(* IEC 61131-3 sources: JingjiangArm/moonboxpro_arm_8.4/Application/Application/任务列表/ExtTask/动作处理/预套准, 13 files *)

(* ---- ENUM_MotionStepIDs.st ---- *)
(*@CES
Name=ENUM_MotionStepIDs
Type=Gvl
TypeGuid=2db5746d-d284-4425-9f7f-2663a34b0ebc
Guid=2f95a26a-5938-4297-8364-5fa39176fcfb
HasDeclaration=True
HasImplementation=False
*)
{DECLARATION}

TYPE ENUM_MotionStepIDs : (
	MOTION_STEP_NothingDo						:= -1,(*啥都不做*)
	MOTION_STEP_MotionCtrlModel				:= 9,(*2021.2.21.134018设置运动模式设置|+Liu.yt*)
	MOTION_STEP_ServoOff					:= 10,(*下伺服|*)
	MOTION_STEP_ClrSts						:= 11,(*清错误状态|*)
	MOTION_STEP_ZeroPos						:= 12,(*清位置|*)
	MOTION_STEP_ZeroPos_Again				:= 13,(*2018.9.4.144137\再次清位置|*)
	MOTION_STEP_ServoOn						:= 14,(*上伺服|*)
	MOTION_STEP_PtModeDynamic				:= 15,(*设置动态pt规划|*)
	MOTION_STEP_PtClear						:= 16,(*清除动态ptFIFO|*)
	MOTION_STEP_SetModal0					:= 17,(*2017-09-11 09:14:16| 模态0*)
	MOTION_STEP_SyncAllModal0				:= 18,(*同步所有轴模态|*)
	MOTION_STEP_SetModal1					:= 19,(*2017-09-11 09:14:24| 模态1*)
	MOTION_STEP_SyncAllModal1				:= 20,(*同步所有轴模态|*)
	MOTION_STEP_WaitingModalChanged			:= 21,(*等待模态切换0到1|*)
	MOTION_STEP_PushInitialPTdata			:= 22,(*压入初始的几段PT数据*)
	MOTION_STEP_WritePT						:= 23,(*写pt*)
	MOTION_STEP_CheckPTPrf					:= 24,(*检查pt规划器*)
	MOTION_STEP_SetTpid						:= 25,(*设置前馈增益|*)
	MOTION_STEP_SetPosErr					:= 26,(*设置位置偏差|*)
	MOTION_STEP_SetEncSns					:= 27,(*编码器反转|*)
	MOTION_STEP_CheckAllServoSts			:= 28,(*检查所有上伺服的状态|*)
	MOTION_STEP_WillLeaveWritePT			:= 29,(*将要离开PT写操作|2019.11.29.143804_*)
	MOTION_STEP_MULTI_GTCMD					:= 30,(*多个指令同时执行标志@单运行功能使用|点了按钮响应太慢了*)
	MOTION_STEP_ErrorOccured				:= 110(*错误发生*)
);
END_TYPE
{IMPLEMENTATION}

(* ---- KS_CalcCircleTangentDistance.st ---- *)
(*@CES
Name=KS_CalcCircleTangentDistance
Type=FunctionBlock
TypeGuid=6f9dac99-8de1-4efc-8465-68ac443b7d08
Guid=1060efe6-291c-4829-ad87-f7b1dbfd88c0
HasDeclaration=True
HasImplementation=True
*)
{DECLARATION}
FUNCTION KS_CalcCircleTangentDistance : LREAL(*计算两个圆的切线距离|*)
VAR_INPUT
	i_lrX_Circle0							: LREAL;(*圆1的圆心坐标x|*)
	i_lrY_Circle0							: LREAL;(*圆1的圆心坐标y|*)
	i_lrDiam_Circle0						: LREAL;(*圆1的直径|*)
	i_lrX_Circle1							: LREAL;(*圆2的圆心坐标x|*)
	i_lrY_Circle1							: LREAL;(*圆2的圆心坐标y|*)
	i_lrDiam_Circle1						: LREAL;(*圆2的直径|*)
	i_xAtSameSide							: BOOL;(*TRUE表示圆是在切线的同一边(外公切)|FALSE表示分别在切线的两边(内公切)|*)
END_VAR
VAR
	lrN										: LREAL;
	lrResult								: LREAL;
	lrCenterDistance						: LREAL;(*两个圆的圆心距|*)
END_VAR
{IMPLEMENTATION}
lrResult:= 0;

(*
/.圆心距|
/.直角三角形的斜边|
/.*)
lrCenterDistance:= SQRT((i_lrX_Circle0-i_lrX_Circle1)*(i_lrX_Circle0-i_lrX_Circle1)+(i_lrY_Circle0-i_lrY_Circle1)*(i_lrY_Circle0-i_lrY_Circle1));
IF i_xAtSameSide THEN
	(*
	/.外公切|
	/.外公切线的长=根号下[圆心距的平方-（大圆半径减小圆半径）的平方]|
	/.*)
	lrN:= (lrCenterDistance*lrCenterDistance)-(((i_lrDiam_Circle0-i_lrDiam_Circle1)/2)*((i_lrDiam_Circle0-i_lrDiam_Circle1)/2));
	IF lrN<0 THEN
		;
	ELSE
		lrResult:= SQRT(lrN);
	END_IF
ELSE
	(*
	/.内公切|
	/.内公切线的长=根号下[圆心距的平方-（大圆半径加小圆半径）的平方]|
	/.*)
	lrN:= (lrCenterDistance*lrCenterDistance)-(((i_lrDiam_Circle0+i_lrDiam_Circle1)/2)*((i_lrDiam_Circle0+i_lrDiam_Circle1)/2));
	IF lrN<0 THEN
		;
	ELSE
		lrResult:= SQRT(lrN);
	END_IF
END_IF
KS_CalcCircleTangentDistance:= lrResult;

(* ---- KS_CalcForPreRegister.st ---- *)
(*@CES
Name=KS_CalcForPreRegister
Type=FunctionBlock
TypeGuid=6f9dac99-8de1-4efc-8465-68ac443b7d08
Guid=6960c73a-5817-444f-97ca-275637423b82
HasDeclaration=True
HasImplementation=True
*)
{DECLARATION}
FUNCTION KS_CalcForPreRegister : WORD(*高8位返回轴号,低8位返回错误*)
(*2023.11.27.104852 欧诺预套准结构同步*)
(*2024.7.11.160354 机组间料长增加翻料架@一般一台机器只有一个翻料架|不支持2个以上翻料架*)
(*那个翻料架应该在当前色和前一色之间*)
(*2024.8.2.173238 调整翻料架料长计算方式*)
VAR_INPUT
	i_iMechanicalType: INT; (*结构类型*)
	i_iGrpAxisNum_Pu: INT; (*色组轴数量*)
	i_aiGrpAxisList: ARRAY [1..MAX_UNIT_NUM] OF INT; (*系内所有轴的列表*)
	i_pstStSysParam: POINTER TO StSysParam;
	i_pastStMechanicalParamBuf: POINTER TO ARRAY [1..5] OF StMechanicalParamBuf; (*机械参数区域*)
	i_iGrpId:INT;(*2024.7.11.164625 输入系id*)
	i_xFilpSwitch:BOOL;(*翻转架开关*)
END_VAR
VAR
	iN: INT;
	iAxisId: INT;

	(*摆臂式机械结构*)
	pstStMechanicalParam_01: POINTER TO StMechanicalParam_01;
	pstStMechanicalParam_03: POINTER TO StMechanicalParam_03;
	pstStMechanicalParam_05: POINTER TO StMechanicalParam_05; (*欧诺直压式结构|2023.07.10.142011*)
	x2,y2: LREAL;
	x4,y4: LREAL;
	lrLCTD1,lrLCTD2,lrLCTD3: LREAL;
	lrVar1,lrVar2,lrVar3,lrVar4: LREAL;
	lrLCirDis_pt1pt3: LREAL; (*pt1到pt3的圆心距*)
	lrLCirDis_pt2pt4: LREAL;
	lrLCirDis_pt2pt5: LREAL;
	lrLCirDis_pt2pt6: LREAL;
	lrLCirDis_pt4pt5: LREAL;
	lrLCirDis_pt4pt6: LREAL;
	lrAng_theta1: LREAL;
	lrAng_q,lrAng_q0: LREAL;
	lrAng_q2: LREAL;
	lrArc_pt5,lrArc_pt4,lrArc_pt2,lrArc_pt6: LREAL;
	lrAng_alpha,lrAng_beta,lrAng_theta,lrAng_delta: LREAL;

	alrConstantLength:ARRAY [1..MAX_UNIT_NUM] OF  LREAL;(*可变料长数组*)
	(*直压式结构*)
	pstStMechanicalParam_02: POINTER TO StMechanicalParam_02; (*机械结构2*)
	lrTotalLength:LREAL;(*总料长*)
	wResult:WORD;
	//pstStAxisParam: POINTER TO StAxisParam;

	lrX_PressRoller: LREAL;
	lrY_PressRoller: LREAL;
	lrLCirDis_pt5ptR: LREAL;
	lrLCirDis_pt6ptR: LREAL;
	lrLCirDis_pt5pt6: LREAL;
	lrAng_65R: LREAL;
	lrAng_5R6: LREAL;
	lrAng_AlphaB: LREAL;
	lrAng_AlphaC: LREAL;
	lrAng_AlphaH: LREAL;
	lrAng_AlphaK: LREAL;
	lrAng_GammaA: LREAL;
	lrAng_GammaB: LREAL;
	lrArc_3: LREAL;
	lrArc_1: LREAL;
	lrArc_2: LREAL;
	X_OnRubberROller: BOOL;
	XH1_Flag: BOOL;		(*胶辊安装在孔H1*)
	XH2_Flag: BOOL;
	lrLCirDis_pt3pt5: LREAL;
	IrO3M: LREAL;
	lrLCirDis_pt2pt3: LREAL;
	IrAngle_O3O2U: LREAL;
	IrAngle_O4O2V: LREAL;
	IrAngle_O3O2O4: LREAL;
	IrAngle_O2O3O5: LREAL;
	IrAngle_O2O3I: LREAL;
	IrAngle_HO3M: LREAL;
	IrAngle_O2O4O6: LREAL;
	IrAngle_O2O4P: LREAL;
	IrAngle_O6O4N: LREAL;
	IrAngle_HO3I: LREAL;
	IrAngle_NO4Q: LREAL;
	IrAngle_WO5S: LREAL;
	IrAngle_ZO5W: LREAL;
	IrArc_UV: LREAL;
	IrArc_HI: LREAL;
	IrArc_NQ: LREAL;
	IrArc_WS: LREAL;
	IrIU: LREAL;
	IrQV: LREAL;
	IrHS: LREAL;
	IrNT: LREAL;
	lrAng_56R:LREAL;
	lrLCirDis_pt3pt6:LREAL;
	IrAngle_UO2V:LREAL;
	IrAngle_O4O3O5:LREAL;
	IrAngle_O3O4O6: LREAL;
	lrLCirDis_pt3pt4: LREAL;
	IrHM: LREAL;
(*2023.07.10.142055|欧诺直压式*)
	lrLCirDis_pt1pt2_LZY : LREAL;
	lrLCirDis_pt2pt3_LZY : LREAL;
	lrLCirDis_pt3pt4_LZY : LREAL;
	lrLCirDis_pt4pt5_LZY : LREAL;
	lrLCirDis_pt5pt6_LZY : LREAL;
	lrLCirDis_pt1pt3_LZY: LREAL;	(*  *)
	lrLCirDis_pt2pt4_LZY: LREAL;	(*  *)
	lrLCirDis_pt3pt5_LZY : LREAL;
	lrLCirDis_pt4pt6_LZY : LREAL;

	lrLCTD1_LZY : LREAL;
	lrLCTD2_LZY : LREAL;
	lrLCTD3_LZY : LREAL;
	lrLCTD4_LZY : LREAL;
	lrLCTD5_LZY : LREAL;
	lrWL1 :LREAL;
	lrWL2 :LREAL;
	lrWL3 :LREAL;
	lrWL4 :LREAL;

	lrWR1 :LREAL;
	lrWR2 :LREAL;
	lrWR3 :LREAL;
	lrWR4 :LREAL;

	lrWU1 :LREAL;
	lrWU2 :LREAL;
	lrWU3 :LREAL;
	lrWU4 :LREAL;
	lrArc1 : LREAL;(*弧长*)
	lrArc2 : LREAL;
	lrArc3 : LREAL;
	lrArc4 : LREAL;
(*2023.11.17.102855*)
	rY3_LD:REAL;

	iError:INT;
	rCentre1_2: REAL; (*棍1和棍2中心的距离*)
	rCentre2_3: REAL;
	rCentre3_4: REAL;
	rCentre1_3: REAL;
	rCentre1_4: REAL;
	rCentre2_4: REAL;
	rCentre3_6: REAL;
	rCentre4_6: REAL;
	rlength2_3: REAL; (*棍2和棍3中心之间的距离,固定不变的*)
	rArcLength2: REAL;  (*棍2上的料长、棍2的弧长*)
	rArcLength3: REAL;
	rArcLength4: REAL;
	rradian_a1: REAL; (*棍1中心和上切点相连的直线与棍1、2中心连线的夹角对应的弧度*)
	rradian_a2: REAL; (*棍1、2中心相连的直线与棍2、3中心相连的直线的夹角对应的弧度*)
	rradian_a3: REAL; (*棍2下切点与棍3左切点相连的直线与棍2、3中心相连的直线的夹角对应的弧度*)
	rradian_a4: REAL;
	rradian_b1: REAL; (*棍3中心与左切点相连的直线与棍2、3中心连线的夹角对应的弧度*)
	rradian_b2: REAL; (*棍2、3中心相连的直线与棍3、4中心相连的直线的夹角对应的弧度*)
	rradian_b3: REAL; (*棍3右切点与棍4下切点相连的直线与棍3、4中心相连的直线的夹角对应的弧度*)
	rradian_c1: REAL; (*棍3右切点与棍4下切点相连的直线与棍3、4中心连线的夹角对应的弧度*)
	rradian_c2: REAL; (*棍3、4中心相连的直线与棍4、6中心相连的直线的夹角对应的弧度*)
	rradian_c3: REAL; (*棍4上切点与棍6下切点相连的直线与棍4、6中心相连的直线的夹角对应的弧度*)
	rradian_c4: REAL;
	rlengthI: REAL;       (*棍1和2间的料长*)

	rlengthII: REAL;      (*棍2和3间的料长*)
	rlengthIII: REAL;	  (*棍3和4间的料长*)
	rLrength4_6: REAL; (*棍4和棍6之间的料长*)
	rTotallength: REAL;   (*总可变料长*)
	rlengthI1: REAL;

	rradian_d1: REAL; (*棍1、2中心相连的直线与棍1的Y1之间的夹角所对应的弧度------2022.10.25.155501*)
	rradian_d2: REAL; (*棍1、2中心相连的直线与棍1中心和下切点相连的直线夹角对应的弧度*)
	rlengthI2: REAL;  (*棍1下切点与棍2中心之间的距离-------2022.10.25.155433*)
	rArcLength1: REAL;  (*棍1上的料长、棍1的弧长--------2022.10.25.155406*)

	//2025.12.24.133817 | + | 秦华程序增加结构6
	pstStUnitParam_Save: POINTER TO StUnitParam_Save;
	pstStUnitParam_UnSave: POINTER TO StUnitParam_UnSave;
	iUnitValid : INT;
	lrTemp_Qinhua : LREAL;
	lrPreReg_Len_V : LREAL;
	xUnitValid : BOOL;

	//品字形 2026.03.10.113914 Hou.N
	rPrRadius:REAL;
	rBrRadius:REAL;
	rHypotenuse:REAL;
	alrAngle_Br: ARRAY [1..MAX_UNIT_NUM] OF  REAL;//底辊压印点和水平的夹角,以水平为基准点
	alrArc_length_Br:ARRAY [1..MAX_UNIT_NUM] OF  REAL;
	lrTemp: LREAL;

	(*2026.08.27.095609*)
	(*欧诺预套准*)
	rPlateR:REAL;(*[AI修改20260827]版辊半径|由本轴rGirth_PrnRoller/π/2推算,替代已删除的rD0/2*)
	rY3:REAL;(*[AI修改20260829]辊3辊心高=动态|Y0+版半径+D3/2,随版径浮动*)
	rL2_3:REAL;(*[AI修改20260829]辊2-3垂直中心距=动态派生|rY2-rY3|原为静态结构体字段*)
	rd1:REAL;(*D1与D2的圆心距*)
	rd2:REAL;(*D2与D3的圆心距*)
	rd3:REAL;(*D3与D4的圆心距*)
	rd4:REAL;(*D1与D3的圆心距*)
	rd5:REAL;(*D2与D4的圆心距*)
	rCenter_To_tangent1:REAL;(*D1圆心与D2切点的距离*)
	rCenter_To_tangent2:REAL;(*D3圆心与D2切点的距离*)
	rCenter_To_tangent3:REAL;(*D2圆心与D3切点的距离*)
	rCenter_To_tangent4:REAL;(*D4圆心与D3切点的距离*)
	rLength1:REAL;(*D1与D2之间料长*)
	rArcLen1:REAL;(*D2辊上的料长-弧长*)
	rLength2:REAL;(*D2与D3之间料长*)
	rArcLen2:REAL;(*D3辊上的料长-弧长*)
	rLength3:REAL;(*D3与D4之间料长*)
	rArc1:REAL;(*角1对应的弧长1*)
	rArc2:REAL;(*角2对应的弧长2*)
	rArc3:REAL;(*角3对应的弧长3*)
	rArc5:REAL;(*角5对应的弧长5*)
	rArc6:REAL;(*角6对应的弧长6*)
	rArc7:REAL;(*角7对应的弧长7*)
	rAngle1:REAL;(*角1*)
	rAngle2:REAL;(*角2*)
	rAngle3:REAL;(*角3*)
	rAngle4:REAL;(*角4-D2所求弧面料长对应的角*)
	rAngle5:REAL;(*角5*)
	rAngle6:REAL;(*角6*)
	rAngle7:REAL;(*角7*)
	rAngle8:REAL;(*角8-D3所求弧面料长对应的角*)

END_VAR

{IMPLEMENTATION}
wResult:= 0;
IF i_pstStSysParam<>0 AND
	i_pastStMechanicalParamBuf<>0 AND
	(i_iGrpAxisNum_Pu>=1 AND i_iGrpAxisNum_Pu<=MAX_UNIT_NUM) AND
	(i_iGrpId=1 OR i_iGrpId=2 ) THEN
	CASE i_iMechanicalType OF
	1: (*摆臂机械结构*)
		pstStMechanicalParam_01:= ADR(i_pastStMechanicalParamBuf^[1].abyBuf);
		IF pstStMechanicalParam_01^.lrX1<0.1 OR pstStMechanicalParam_01^.lry1<0.1 OR  pstStMechanicalParam_01^.lrx3<0.1
			OR  pstStMechanicalParam_01^.lry3<0.1 OR  pstStMechanicalParam_01^.lrx5<0.1 OR  pstStMechanicalParam_01^.lry5<0.1
			OR  pstStMechanicalParam_01^.lrx6<0.1  OR  pstStMechanicalParam_01^.lry6<0.1 THEN
			wResult:=16#FF01;
			RETURN;
		END_IF

		FOR iN:=1 TO i_iGrpAxisNum_Pu BY 1 DO
			iAxisId:= i_aiGrpAxisList[iN];
			lrVar1:= (pstStMechanicalParam_01^.lrX1 - pstStMechanicalParam_01^.lrX3);
			lrVar2:= (pstStMechanicalParam_01^.lrY1 - pstStMechanicalParam_01^.lrY3);
			lrLCirDis_pt1pt3:= SQRT(lrVar1*lrVar1 + lrVar2*lrVar2);
			lrVar1:= lrLCirDis_pt1pt3;
			lrVar2:= (pstStMechanicalParam_01^.lrL2);
			lrVar3:= ((i_pstStSysParam^.astStUnitParam_Save[iAxisId].rGirth_PrnRoller)/gc_lrPI + (pstStMechanicalParam_01^.lrDR))/2;

			IF lrVar1=0 OR lrVar2=0 OR lrLCirDis_pt1pt3=0 THEN
				wResult:=SHL(INT_TO_WORD(iN),8)+16#0002;
				EXIT;
			END_IF

			lrVar4:= (lrVar1*lrVar1+lrVar2*lrVar2-lrVar3*lrVar3) / (2*lrVar1*lrVar2);
			IF  ABS(lrVar4)>1 THEN
				wResult:=SHL(INT_TO_WORD(iN),8)+16#0003;
				EXIT;
			END_IF

			lrAng_q:= ACOS( (lrVar1*lrVar1+lrVar2*lrVar2-lrVar3*lrVar3) / (2*lrVar1*lrVar2) ); (*余弦定理*)

			lrVar4:=(pstStMechanicalParam_01^.lrY3-pstStMechanicalParam_01^.lrY1) / lrLCirDis_pt1pt3 ;
			IF  ABS(lrVar4)>1 THEN
				wResult:=SHL(INT_TO_WORD(iN),8)+16#0004;
				EXIT;
			END_IF
			lrAng_q0:= ASIN( (pstStMechanicalParam_01^.lrY3-pstStMechanicalParam_01^.lrY1) / lrLCirDis_pt1pt3 );
			lrAng_theta1:= lrAng_q - lrAng_q0; (*如果pt3高过pt2,则包角相减<0，并不会影响到pt2的计算*)

			x2:= pstStMechanicalParam_01^.lrX3 + (pstStMechanicalParam_01^.lrL2)*COS(lrAng_theta1);
			y2:= pstStMechanicalParam_01^.lrY3 + (pstStMechanicalParam_01^.lrL2)*SIN(lrAng_theta1);

			lrAng_q2:= gc_lrPI - (pstStMechanicalParam_01^.lrA)*(gc_lrPI/180.0) - lrAng_theta1;

			x4:= pstStMechanicalParam_01^.lrX3-(pstStMechanicalParam_01^.lrL1)*COS(lrAng_q2);
			y4:= pstStMechanicalParam_01^.lrY3+(pstStMechanicalParam_01^.lrL1)*SIN(lrAng_q2);

	        (*切线段长度*)
			lrLCTD1:= KS_CalcCircleTangentDistance(
				pstStMechanicalParam_01^.lrX5, pstStMechanicalParam_01^.lrY5, pstStMechanicalParam_01^.lrD1,
				x4, y4, pstStMechanicalParam_01^.lrD2,
				FALSE);

			lrLCTD2:= KS_CalcCircleTangentDistance(
				x4, y4, pstStMechanicalParam_01^.lrD2,
				x2, y2, pstStMechanicalParam_01^.lrDR,
				TRUE);

			lrLCTD3:= KS_CalcCircleTangentDistance(
				x2, y2, pstStMechanicalParam_01^.lrDR,
				pstStMechanicalParam_01^.lrX6, pstStMechanicalParam_01^.lrY6, pstStMechanicalParam_01^.lrD3,
				TRUE);

	        (*临近的圆心距*)
			lrVar1:= x2-x4;
	        lrVar2:= y2-y4;
	        lrLCirDis_pt2pt4:= SQRT( lrVar1*lrVar1 + lrVar2*lrVar2 );

	        lrVar1:= x2 - (pstStMechanicalParam_01^.lrX5);
	        lrVar2:= y2 - (pstStMechanicalParam_01^.lrY5);
	        lrLCirDis_pt2pt5:= SQRT( lrVar1*lrVar1 + lrVar2*lrVar2 );

	        lrVar1:= x2 - (pstStMechanicalParam_01^.lrX6);
	        lrVar2:= y2 - (pstStMechanicalParam_01^.lrY6);
	        lrLCirDis_pt2pt6:= SQRT( lrVar1*lrVar1 + lrVar2*lrVar2 );

	        lrVar1:= x4 - (pstStMechanicalParam_01^.lrX6);
	        lrVar2:= y4 - (pstStMechanicalParam_01^.lrY6);
	        lrLCirDis_pt4pt6:= SQRT( lrVar1*lrVar1 + lrVar2*lrVar2 );

	        lrVar1:= x4 - (pstStMechanicalParam_01^.lrX5);
	        lrVar2:= y4 - (pstStMechanicalParam_01^.lrY5);
	        lrLCirDis_pt4pt5:= SQRT( lrVar1*lrVar1 + lrVar2*lrVar2 );

			IF lrLCirDis_pt4pt5=0 OR
				lrLCirDis_pt2pt4=0 OR
				lrLCirDis_pt2pt6=0 THEN (*2017-09-05 11:26:10|*)
				wResult:=SHL(INT_TO_WORD(iN),8)+16#0005;
				EXIT;
			END_IF
	        lrVar1:= (pstStMechanicalParam_01^.lrX5)-x4;
	        lrVar2:= ((pstStMechanicalParam_01^.lrD1) + (pstStMechanicalParam_01^.lrD2))/2.0;
			lrVar4:=lrVar1/lrLCirDis_pt4pt5;
			IF  ABS(lrVar4)>1 THEN
				wResult:=SHL(INT_TO_WORD(iN),8)+16#0006;
				EXIT;
			END_IF

			lrVar4:=lrVar2/lrLCirDis_pt4pt5;
			IF  ABS(lrVar4)>1 THEN
				wResult:=SHL(INT_TO_WORD(iN),8)+16#0007;
				EXIT;
			END_IF
	        lrAng_alpha:= ASIN(lrVar1/lrLCirDis_pt4pt5) + ASIN(lrVar2/lrLCirDis_pt4pt5); (*pt5弧角*)

	        lrVar1:= ((pstStMechanicalParam_01^.lrDR) - (pstStMechanicalParam_01^.lrD2))/2.0;
	        lrVar2:= x2-x4;
			lrVar4:=lrVar1/lrLCirDis_pt2pt4;
			IF  ABS(lrVar4)>1 THEN
				wResult:=SHL(INT_TO_WORD(iN),8)+16#0008;
				EXIT;
			END_IF

			lrVar4:=lrVar2/lrLCirDis_pt2pt4;
			IF  ABS(lrVar4)>1 THEN
				wResult:=SHL(INT_TO_WORD(iN),8)+16#0009;
				EXIT;
			END_IF
	        lrAng_beta:= ACOS(lrVar1/lrLCirDis_pt2pt4) - ACOS(lrVar2/lrLCirDis_pt2pt4); (*与alpha合并构成pt4弧角*)

	        lrVar1:= ((pstStMechanicalParam_01^.lrDR) - (pstStMechanicalParam_01^.lrD3))/2.0;
	        lrVar2:= (pstStMechanicalParam_01^.lrX6) - x2;
			lrVar4:=lrVar1/lrLCirDis_pt2pt6;
			IF  ABS(lrVar4)>1 THEN
				wResult:=SHL(INT_TO_WORD(iN),8)+16#000A;
				EXIT;
			END_IF

			lrVar4:=lrVar2/lrLCirDis_pt2pt6;
			IF  ABS(lrVar4)>1 THEN
				wResult:=SHL(INT_TO_WORD(iN),8)+16#000B;
				EXIT;
			END_IF
	        lrAng_delta:= ACOS(lrVar1/lrLCirDis_pt2pt6) - ACOS(lrVar2/lrLCirDis_pt2pt6); (*pt6弧角*)

	        lrAng_theta:= gc_lrPI - lrAng_beta - lrAng_delta; (*压辊弧角*)

	        lrArc_pt5:= ((pstStMechanicalParam_01^.lrD1)/2)*lrAng_alpha;
	        lrArc_pt4:= ((pstStMechanicalParam_01^.lrD2)/2)*(lrAng_alpha+lrAng_beta);
	        lrArc_pt2:= ((pstStMechanicalParam_01^.lrDR)/2)*lrAng_theta;
	        lrArc_pt6:= ((pstStMechanicalParam_01^.lrD3)/2)*lrAng_delta;
			alrConstantLength[iN]:=lrArc_pt5+lrLCTD1+lrArc_pt4+lrLCTD2+lrArc_pt2+lrLCTD3+lrArc_pt6;
			lrTotalLength:=alrConstantLength[iN]+i_pstStSysParam^.astStUnitParam_Save[iAxisId].lrPreReg_ConstVal;
			(*2024.7.11.164906+*)

			IF i_xFilpSwitch THEN(*翻转架开关打开了|就把翻料架的料长加进去@一般一台机器只有一个翻料架*)
				IF i_pstStSysParam^.astStGrpParam_Save[i_iGrpId].byTurnOverAxisId=0 THEN(*=0|那个轴有翻料架值就直接累加*)
					lrTotalLength:=lrTotalLength+i_pstStSysParam^.astStUnitParam_Save[iAxisId].uiTurnOverFilmLenth;
				ELSE
					IF i_pstStSysParam^.astStGrpParam_Save[i_iGrpId].byTurnOverAxisId=iAxisId THEN(*就是输入的轴id@累加该轴的翻料架长度*)
						lrTotalLength:=lrTotalLength+i_pstStSysParam^.astStUnitParam_Save[iAxisId].uiTurnOverFilmLenth;
					END_IF
				END_IF
			END_IF

			IF iN=1 THEN
				lrTotalLength:=0;
				i_pstStSysParam^.astStUnitParam_Save[iAxisId].lrPreReg_Length_V:=0;
				i_pstStSysParam^.astStUnitParam_Save[iAxisId].lrFilmLengthFromPrevUnit:=lrTotalLength;
			ELSE
				i_pstStSysParam^.astStUnitParam_Save[iAxisId].lrFilmLengthFromPrevUnit:=lrTotalLength;
				i_pstStSysParam^.astStUnitParam_Save[iAxisId].lrPreReg_Length_V:= KS_LREAL_MOD(lrTotalLength, i_pstStSysParam^.astStUnitParam_Save[iAxisId].rGirth_PrnRoller); (* 当前色预套准计算的值 *)
				i_pstStSysParam^.astStUnitParam_Save[iAxisId].lrPreReg_Length_V:=
									(i_pstStSysParam^.astStUnitParam_Save[iAxisId].rGirth_PrnRoller-i_pstStSysParam^.astStUnitParam_Save[iAxisId].lrPreReg_Length_V) + (* 版向走料方向单方向运动的是余数部分 *)
									i_pstStSysParam^.astStUnitParam_Save[iAxisId].lrPreReg_Adjust + (* 输入的修正值 *)
									i_pstStSysParam^.astStUnitParam_Save[i_aiGrpAxisList[iN-1]].lrPreReg_Length_V; (* 前一色已经运动过的量|相当于更新变化后的基准位置 *)

				(* 2020.9.11.152457|防止输入的修正值绝对值超出1个版周 *)
				WHILE i_pstStSysParam^.astStUnitParam_Save[iAxisId].lrPreReg_Length_V<0 DO
					i_pstStSysParam^.astStUnitParam_Save[iAxisId].lrPreReg_Length_V:= i_pstStSysParam^.astStUnitParam_Save[iAxisId].lrPreReg_Length_V+i_pstStSysParam^.astStUnitParam_Save[iAxisId].rGirth_PrnRoller;
				END_WHILE
				WHILE i_pstStSysParam^.astStUnitParam_Save[iAxisId].lrPreReg_Length_V>i_pstStSysParam^.astStUnitParam_Save[iAxisId].rGirth_PrnRoller DO
					i_pstStSysParam^.astStUnitParam_Save[iAxisId].lrPreReg_Length_V:= i_pstStSysParam^.astStUnitParam_Save[iAxisId].lrPreReg_Length_V-i_pstStSysParam^.astStUnitParam_Save[iAxisId].rGirth_PrnRoller;
				END_WHILE

			END_IF
		END_FOR
	2: (*直压式结构*)
		pstStMechanicalParam_02:= ADR(i_pastStMechanicalParamBuf^[2].abyBuf);
		IF pstStMechanicalParam_02^.lrX1<0.1 OR pstStMechanicalParam_02^.lry1<0.1 OR  pstStMechanicalParam_02^.lrx5<0.1
			OR  pstStMechanicalParam_02^.lry5<0.1 OR  pstStMechanicalParam_02^.lrx6<0.1  OR  pstStMechanicalParam_02^.lry6<0.1 THEN
			wResult:=16#FF01;
			RETURN;
		END_IF
		FOR iN:=1 TO i_iGrpAxisNum_Pu BY 1 DO
			iAxisId:= i_aiGrpAxisList[iN];
			lrX_PressRoller:=pstStMechanicalParam_02^.lrX1;
			lrY_PressRoller:= pstStMechanicalParam_02^.lry1-((i_pstStSysParam^.astStUnitParam_Save[iAxisId].rGirth_PrnRoller)/gc_lrPI+pstStMechanicalParam_02^.lrDR)/2.0;
			(*算出左边导向辊和胶辊之间的圆心距离*)
			lrVar1:= (lrX_PressRoller-pstStMechanicalParam_02^.lrx5);
			lrVar2:= (lrY_PressRoller-pstStMechanicalParam_02^.lrY5);
			lrLCirDis_pt5ptR:= SQRT(lrVar1*lrVar1 + lrVar2*lrVar2);
			(*算出右边导向辊和胶辊之间的圆心距离*)
			lrVar1:= (pstStMechanicalParam_02^.lrx6-lrX_PressRoller);
			lrVar2:= (pstStMechanicalParam_02^.lry6-lrY_PressRoller);
			lrLCirDis_pt6ptR:= SQRT(lrVar1*lrVar1 + lrVar2*lrVar2);
			(*算出x5,y5和x6,y6之间的圆心距离*)
			lrVar1:= pstStMechanicalParam_02^.lrx6-pstStMechanicalParam_02^.lrx5;
			lrVar2:= pstStMechanicalParam_02^.lrY6-pstStMechanicalParam_02^.lrY5;
			lrLCirDis_pt5pt6:= SQRT(lrVar1*lrVar1 + lrVar2*lrVar2);
			IF NOT (lrLCirDis_pt5ptR<>0 AND lrLCirDis_pt6ptR<>0) THEN(*分母不能为0*)
				wResult:=SHL(INT_TO_WORD(iN),8)+16#0002;
				EXIT;
			END_IF
			IF ABS((lrLCirDis_pt5ptR*lrLCirDis_pt5ptR + lrLCirDis_pt6ptR*lrLCirDis_pt6ptR - lrLCirDis_pt5pt6*lrLCirDis_pt5pt6) / (2*lrLCirDis_pt5ptR*lrLCirDis_pt6ptR)) > 1 THEN (*余弦值域必须有效*)
				wResult:=SHL(INT_TO_WORD(iN),8)+16#0003;
				EXIT;
			END_IF
			(*算出x5,y5|胶辊|x6,y6的夹角*)
			(*余弦定理| cos(abc)=(a2+b2-c2)/2ab*)
			lrAng_5R6:= ACOS((lrLCirDis_pt5ptR*lrLCirDis_pt5ptR + lrLCirDis_pt6ptR*lrLCirDis_pt6ptR - lrLCirDis_pt5pt6*lrLCirDis_pt5pt6) / (2*lrLCirDis_pt5ptR*lrLCirDis_pt6ptR));
			(*两段切线|都是外切*)
			(*左边导向辊到压辊之间的外切线距离*)
			lrLCTD1:= KS_CalcCircleTangentDistance(
				pstStMechanicalParam_02^.lrx5, pstStMechanicalParam_02^.lrY5, pstStMechanicalParam_02^.lrD1,
				lrX_PressRoller, lrY_PressRoller, pstStMechanicalParam_02^.lrDR,
				FALSE);

			lrLCTD2:= KS_CalcCircleTangentDistance(
				pstStMechanicalParam_02^.lrX6, pstStMechanicalParam_02^.lrY6, pstStMechanicalParam_02^.lrD3,
				lrX_PressRoller, lrY_PressRoller, pstStMechanicalParam_02^.lrDR,
				FALSE);
			IF NOT (lrLCirDis_pt5pt6<>0 AND lrLCirDis_pt5ptR<>0) THEN(*分母不能0*)
				wResult:=SHL(INT_TO_WORD(iN),8)+16#0004;
				EXIT;
			END_IF
			IF ABS((lrLCirDis_pt5ptR*lrLCirDis_pt5ptR + lrLCirDis_pt5pt6*lrLCirDis_pt5pt6 - lrLCirDis_pt6ptR*lrLCirDis_pt6ptR) / (2*lrLCirDis_pt5pt6*lrLCirDis_pt5ptR)) > 1 THEN(*余弦值域必须有效*)
				wResult:=SHL(INT_TO_WORD(iN),8)+16#0005;
				EXIT;
			END_IF
			(*将来要用来计算弧长的几个角度*)
			lrAng_65R:= ACOS((lrLCirDis_pt5ptR*lrLCirDis_pt5ptR + lrLCirDis_pt5pt6*lrLCirDis_pt5pt6 - lrLCirDis_pt6ptR*lrLCirDis_pt6ptR) / (2*lrLCirDis_pt5pt6*lrLCirDis_pt5ptR));
			lrAng_56R:= gc_lrPI-lrAng_65R-lrAng_5R6;
			IF ABS((lrX_PressRoller-pstStMechanicalParam_02^.lrx5)/lrLCirDis_pt5ptR)>1 THEN(*asin()值域必须检查*)
				wResult:=SHL(INT_TO_WORD(iN),8)+16#0006;
				EXIT;
			END_IF
			lrAng_AlphaB:= ASIN((lrX_PressRoller-pstStMechanicalParam_02^.lrx5)/lrLCirDis_pt5ptR);

			IF ABS(lrLCTD1/lrLCirDis_pt5ptR)>1 THEN(*acos()值域必须检查*)
				wResult:=SHL(INT_TO_WORD(iN),8)+16#0007;
				EXIT;
			END_IF
			lrAng_AlphaC:= ACOS(lrLCTD1/lrLCirDis_pt5ptR);
			lrAng_GammaA:= lrAng_AlphaB-lrAng_AlphaC; (*A点开始的弧角*)
			IF ABS(lrLCTD2/lrLCirDis_pt6ptR)>1 THEN(*asin()值域必须有效*)
				wResult:=SHL(INT_TO_WORD(iN),8)+16#0008;
				EXIT;
			END_IF
			lrAng_Beta:= 2*gc_lrPI - lrAng_5R6 - ASIN(lrLCTD1/lrLCirDis_pt5ptR) - ASIN(lrLCTD2/lrLCirDis_pt6ptR);
			IF ABS((pstStMechanicalParam_02^.lrX6-lrX_PressRoller)/lrLCirDis_pt6ptR)>1 THEN(*asin()值域检查*)
				wResult:=SHL(INT_TO_WORD(iN),8)+16#0009;
				EXIT;
			END_IF
			lrAng_AlphaH:= ASIN((pstStMechanicalParam_02^.lrX6-lrX_PressRoller)/lrLCirDis_pt6ptR);

			IF ABS(lrLCTD2/lrLCirDis_pt6ptR)>1 THEN(*acos()值域检查*)
				wResult:=SHL(INT_TO_WORD(iN),8)+16#000A;
				EXIT;
			END_IF
			lrAng_AlphaK:= ACOS(lrLCTD2/lrLCirDis_pt6ptR);
			lrAng_GammaB:= lrAng_AlphaH-lrAng_AlphaK;
			(*弧长A点在x5,y5上的弧线长度*)
			lrArc_1:= (pstStMechanicalParam_02^.lrD1/2.0)*lrAng_GammaA;

			(*弧长在压辊上的长度*)
			lrArc_2:= (pstStMechanicalParam_02^.lrDR/2.0)*lrAng_Beta;

			(*弧长B点在x6,y6上的弧线长度*)
			lrArc_3:= (pstStMechanicalParam_02^.lrD3/2.0)*lrAng_GammaB;
			alrConstantLength[iN]:= lrArc_1+lrLCTD1+lrArc_2+lrLCTD2+lrArc_3;
			lrTotalLength:=alrConstantLength[iN]+i_pstStSysParam^.astStUnitParam_Save[iAxisId].lrPreReg_ConstVal;
			(*2024.7.11.164906+*)

			IF i_xFilpSwitch THEN(*翻转架开关打开了|就把翻料架的料长加进去@一般一台机器只有一个翻料架*)
				IF i_pstStSysParam^.astStGrpParam_Save[i_iGrpId].byTurnOverAxisId=0 THEN(*=0|那个轴有翻料架值就直接累加*)
					lrTotalLength:=lrTotalLength+i_pstStSysParam^.astStUnitParam_Save[iAxisId].uiTurnOverFilmLenth;
				ELSE
					IF i_pstStSysParam^.astStGrpParam_Save[i_iGrpId].byTurnOverAxisId=iAxisId THEN(*就是输入的轴id@累加该轴的翻料架长度*)
						lrTotalLength:=lrTotalLength+i_pstStSysParam^.astStUnitParam_Save[iAxisId].uiTurnOverFilmLenth;
					END_IF
				END_IF
			END_IF

			IF iN=1 THEN
				lrTotalLength:=0;
				i_pstStSysParam^.astStUnitParam_Save[iAxisId].lrPreReg_Length_V:=0;
				i_pstStSysParam^.astStUnitParam_Save[iAxisId].lrFilmLengthFromPrevUnit:=lrTotalLength;
			ELSE
				i_pstStSysParam^.astStUnitParam_Save[iAxisId].lrFilmLengthFromPrevUnit:=lrTotalLength;
				i_pstStSysParam^.astStUnitParam_Save[iAxisId].lrPreReg_Length_V:= KS_LREAL_MOD(lrTotalLength, i_pstStSysParam^.astStUnitParam_Save[iAxisId].rGirth_PrnRoller);(*当前色预套准计算的值*)
				i_pstStSysParam^.astStUnitParam_Save[iAxisId].lrPreReg_Length_V:=i_pstStSysParam^.astStUnitParam_Save[iAxisId].rGirth_PrnRoller-i_pstStSysParam^.astStUnitParam_Save[iAxisId].lrPreReg_Length_V
									+i_pstStSysParam^.astStUnitParam_Save[iAxisId].lrPreReg_Adjust+i_pstStSysParam^.astStUnitParam_Save[i_aiGrpAxisList[iN-1]].lrPreReg_Length_V;

				(* 2020.9.11.152457|防止输入的修正值绝对值超出1个版周 *)
				WHILE i_pstStSysParam^.astStUnitParam_Save[iAxisId].lrPreReg_Length_V<0 DO
					i_pstStSysParam^.astStUnitParam_Save[iAxisId].lrPreReg_Length_V:= i_pstStSysParam^.astStUnitParam_Save[iAxisId].lrPreReg_Length_V+i_pstStSysParam^.astStUnitParam_Save[iAxisId].rGirth_PrnRoller;
				END_WHILE
				WHILE i_pstStSysParam^.astStUnitParam_Save[iAxisId].lrPreReg_Length_V>i_pstStSysParam^.astStUnitParam_Save[iAxisId].rGirth_PrnRoller DO
					i_pstStSysParam^.astStUnitParam_Save[iAxisId].lrPreReg_Length_V:= i_pstStSysParam^.astStUnitParam_Save[iAxisId].lrPreReg_Length_V-i_pstStSysParam^.astStUnitParam_Save[iAxisId].rGirth_PrnRoller;
				END_WHILE

			END_IF
		END_FOR
	3:(*欧泰直压式*)
		(*M点为圆3和圆5之间圆心距与切线的交点,
		IrHW为圆3和圆5的切线,H为圆3上的切点,W为圆5上的切点;
		IrNT为圆4和圆6的切线,N为圆4上的切点,T为圆6上的切点;
		IrIU为圆3和圆2的切线,I为圆3上的切点,U为圆5上的切点;
		IrQV为圆4和圆2的切线,Q为圆4上的切点,V为圆6上的切点;
		*)
		pstStMechanicalParam_03:= ADR(i_pastStMechanicalParamBuf^[3].abyBuf);
		IF pstStMechanicalParam_03^.lrX1<0.1 OR pstStMechanicalParam_03^.lry1<0.1 OR  pstStMechanicalParam_03^.lrx3<0.1
			OR  pstStMechanicalParam_03^.lrx4<0.1 OR  pstStMechanicalParam_03^.lrx5<0.1 OR  pstStMechanicalParam_03^.lrx6<0.1  OR  pstStMechanicalParam_03^.lry6<0.1 THEN
			wResult:=16#FF01;
			RETURN;
		END_IF
		pstStMechanicalParam_03^.lrX2:=pstStMechanicalParam_03^.lrX1;
		FOR iN:=1 TO i_iGrpAxisNum_Pu BY 1 DO
			iAxisId:= i_aiGrpAxisList[iN];

			pstStMechanicalParam_03^.lrY2:=pstStMechanicalParam_03^.lrY1+0.5*((i_pstStSysParam^.astStUnitParam_Save[iAxisId].rGirth_PrnRoller)/gc_lrPI+pstStMechanicalParam_03^.lrD2);
			IF X_OnRubberROller THEN(*胶辊安装位置确定*)
				pstStMechanicalParam_03^.lrY3:=pstStMechanicalParam_03^.lrY2+pstStMechanicalParam_03^.lrn;
				pstStMechanicalParam_03^.lrY4:=pstStMechanicalParam_03^.lrY2+pstStMechanicalParam_03^.lrm;
				XH1_Flag:=TRUE;
				XH2_Flag:=FALSE;
			ELSE
				XH2_Flag:=TRUE;
				XH1_Flag:=FALSE;
				pstStMechanicalParam_03^.lrY3:=pstStMechanicalParam_03^.lrY2+pstStMechanicalParam_03^.lrn+pstStMechanicalParam_03^.lrH12;
				pstStMechanicalParam_03^.lrY4:=pstStMechanicalParam_03^.lrY2+pstStMechanicalParam_03^.lrm+pstStMechanicalParam_03^.lrH12;
			END_IF
			(*以下为每个圆心之间的距离*)
			lrLCirDis_pt2pt3:=SQRT((pstStMechanicalParam_03^.lrY3-pstStMechanicalParam_03^.lrY2)*(pstStMechanicalParam_03^.lrY3-pstStMechanicalParam_03^.lrY2)
									+(pstStMechanicalParam_03^.lrX3-pstStMechanicalParam_03^.lrX2)*(pstStMechanicalParam_03^.lrX3-pstStMechanicalParam_03^.lrX2));
			lrLCirDis_pt2pt4:=SQRT((pstStMechanicalParam_03^.lrY4-pstStMechanicalParam_03^.lrY2)*(pstStMechanicalParam_03^.lrY4-pstStMechanicalParam_03^.lrY2)
									+(pstStMechanicalParam_03^.lrX4-pstStMechanicalParam_03^.lrX2)*(pstStMechanicalParam_03^.lrX4-pstStMechanicalParam_03^.lrX2));
			lrLCirDis_pt3pt4:=SQRT((pstStMechanicalParam_03^.lrY4-pstStMechanicalParam_03^.lrY3)*(pstStMechanicalParam_03^.lrY4-pstStMechanicalParam_03^.lrY3)
									+(pstStMechanicalParam_03^.lrX4-pstStMechanicalParam_03^.lrX3)*(pstStMechanicalParam_03^.lrX4-pstStMechanicalParam_03^.lrX3));
			lrLCirDis_pt3pt5:=SQRT((pstStMechanicalParam_03^.lrY5-pstStMechanicalParam_03^.lrY3)*(pstStMechanicalParam_03^.lrY5-pstStMechanicalParam_03^.lrY3)
									+(pstStMechanicalParam_03^.lrX5-pstStMechanicalParam_03^.lrX3)*(pstStMechanicalParam_03^.lrX5-pstStMechanicalParam_03^.lrX3));
			lrLCirDis_pt4pt5:=SQRT((pstStMechanicalParam_03^.lrY5-pstStMechanicalParam_03^.lrY4)*(pstStMechanicalParam_03^.lrY5-pstStMechanicalParam_03^.lrY4)
									+(pstStMechanicalParam_03^.lrX5-pstStMechanicalParam_03^.lrX4)*(pstStMechanicalParam_03^.lrX5-pstStMechanicalParam_03^.lrX4));
			lrLCirDis_pt4pt6:=SQRT((pstStMechanicalParam_03^.lrY6-pstStMechanicalParam_03^.lrY4)*(pstStMechanicalParam_03^.lrY6-pstStMechanicalParam_03^.lrY4)
									+(pstStMechanicalParam_03^.lrX6-pstStMechanicalParam_03^.lrX4)*(pstStMechanicalParam_03^.lrX6-pstStMechanicalParam_03^.lrX4));
			lrLCirDis_pt3pt6:=SQRT((pstStMechanicalParam_03^.lrY6-pstStMechanicalParam_03^.lrY3)*(pstStMechanicalParam_03^.lrY6-pstStMechanicalParam_03^.lrY3)
									+(pstStMechanicalParam_03^.lrX6-pstStMechanicalParam_03^.lrX3)*(pstStMechanicalParam_03^.lrX6-pstStMechanicalParam_03^.lrX3));
			lrLCirDis_pt2pt6:=SQRT((pstStMechanicalParam_03^.lrY6-pstStMechanicalParam_03^.lrY2)*(pstStMechanicalParam_03^.lrY6-pstStMechanicalParam_03^.lrY2)
									+(pstStMechanicalParam_03^.lrX2-pstStMechanicalParam_03^.lrX6)*(pstStMechanicalParam_03^.lrX2-pstStMechanicalParam_03^.lrX6));
			lrLCirDis_pt2pt5:=SQRT((pstStMechanicalParam_03^.lrY5-pstStMechanicalParam_03^.lrY2)*(pstStMechanicalParam_03^.lrY5-pstStMechanicalParam_03^.lrY2)
									+(pstStMechanicalParam_03^.lrX2-pstStMechanicalParam_03^.lrX5)*(pstStMechanicalParam_03^.lrX2-pstStMechanicalParam_03^.lrX5));
			(*以下为图中需要用到的直线距离、按标识可找到*)
			IrO3M:=(pstStMechanicalParam_03^.lrD3*lrLCirDis_pt3pt5)/(pstStMechanicalParam_03^.lrD3+pstStMechanicalParam_03^.lrD5);
			IrHM:=SQRT(IrO3M*IrO3M-(pstStMechanicalParam_03^.lrD3*pstStMechanicalParam_03^.lrD3)/4);
			IF lrLCirDis_pt2pt5*IrO3M*lrLCirDis_pt2pt3 * lrLCirDis_pt2pt4 * lrLCirDis_pt3pt4 * lrLCirDis_pt3pt5 * lrLCirDis_pt4pt5 * lrLCirDis_pt4pt6 * lrLCirDis_pt3pt6 * lrLCirDis_pt2pt6=0 THEN(*分母不能为零*)
				wResult:=SHL(INT_TO_WORD(iN),8)+16#0002;
				EXIT;
			END_IF
			(*以下为图中需要用到的角度，通过标注可找到*)
			IrAngle_O3O2U:=ACOS(ABS(pstStMechanicalParam_03^.lrD2-pstStMechanicalParam_03^.lrD3)*0.5/lrLCirDis_pt2pt3);
			IF ABS(ABS(pstStMechanicalParam_03^.lrD2-pstStMechanicalParam_03^.lrD3)*0.5/lrLCirDis_pt2pt3)>1 THEN(*正余弦值域的绝对值必须小于1*)
				wResult:=SHL(INT_TO_WORD(iN),8)+16#0003;
				EXIT;
			END_IF
			IrAngle_O4O2V:=ACOS(ABS(pstStMechanicalParam_03^.lrD2-pstStMechanicalParam_03^.lrD4)*0.5/lrLCirDis_pt2pt4);
			IF ABS(ABS(pstStMechanicalParam_03^.lrD2-pstStMechanicalParam_03^.lrD4)*0.5/lrLCirDis_pt2pt4)>1 THEN
				wResult:=SHL(INT_TO_WORD(iN),8)+16#0004;
				EXIT;
			END_IF
			IrAngle_O3O2O4:=ACOS((lrLCirDis_pt2pt3*lrLCirDis_pt2pt3+lrLCirDis_pt2pt4*lrLCirDis_pt2pt4
													-lrLCirDis_pt3pt4*lrLCirDis_pt3pt4)/(2*lrLCirDis_pt2pt3*lrLCirDis_pt2pt4));
			IF ABS((lrLCirDis_pt2pt3*lrLCirDis_pt2pt3+lrLCirDis_pt2pt4*lrLCirDis_pt2pt4
													-lrLCirDis_pt3pt4*lrLCirDis_pt3pt4)/(2*lrLCirDis_pt2pt3*lrLCirDis_pt2pt4))>1 THEN
				wResult:=SHL(INT_TO_WORD(iN),8)+16#0005;
				EXIT;
			END_IF
			IrAngle_UO2V:=2*gc_lrPI-IrAngle_O3O2U-IrAngle_O4O2V-IrAngle_O3O2O4;(*圆2上需要计算的弧度*)

			IrAngle_O4O3O5:=ACOS((lrLCirDis_pt3pt5*lrLCirDis_pt3pt5+lrLCirDis_pt3pt4*lrLCirDis_pt3pt4-lrLCirDis_pt4pt5*lrLCirDis_pt4pt5)/(2*lrLCirDis_pt3pt4*lrLCirDis_pt3pt5));
			IF ABS((lrLCirDis_pt3pt5*lrLCirDis_pt3pt5+lrLCirDis_pt3pt4*lrLCirDis_pt3pt4-lrLCirDis_pt4pt5*lrLCirDis_pt4pt5)/(2*lrLCirDis_pt3pt4*lrLCirDis_pt3pt5))>1 THEN
				wResult:=SHL(INT_TO_WORD(iN),8)+16#0006;
				EXIT;
			END_IF
			IrAngle_O2O3O5:=ACOS((lrLCirDis_pt2pt3*lrLCirDis_pt2pt3+lrLCirDis_pt3pt5*lrLCirDis_pt3pt5-lrLCirDis_pt2pt5*lrLCirDis_pt2pt5)/(2*lrLCirDis_pt2pt3*lrLCirDis_pt3pt5));
			IF ABS((lrLCirDis_pt2pt3*lrLCirDis_pt2pt3+lrLCirDis_pt3pt5*lrLCirDis_pt3pt5-lrLCirDis_pt2pt5*lrLCirDis_pt2pt5)/(2*lrLCirDis_pt2pt3*lrLCirDis_pt3pt5))>1 THEN
				wResult:=SHL(INT_TO_WORD(iN),8)+16#0007;
				EXIT;
			END_IF
			IrAngle_HO3M:=ACOS(pstStMechanicalParam_03^.lrD3/(2*IrO3M));
			IF ABS(pstStMechanicalParam_03^.lrD3/(2*IrO3M))>1 THEN
				wResult:=SHL(INT_TO_WORD(iN),8)+16#0008;
				EXIT;
			END_IF
			IrAngle_O2O3I:=gc_lrPI-IrAngle_O3O2U;
			IrAngle_HO3I:=2*gc_lrPI-IrAngle_O2O3O5-IrAngle_O2O3I-IrAngle_HO3M;(*圆3上需要计算的弧度*)

			IrAngle_O6O4N:=ACOS((ABS(pstStMechanicalParam_03^.lrD4-pstStMechanicalParam_03^.lrD6))/(2*lrLCirDis_pt4pt6));
			IF ABS((ABS(pstStMechanicalParam_03^.lrD4-pstStMechanicalParam_03^.lrD6))/(2*lrLCirDis_pt4pt6))>1 THEN
				wResult:=SHL(INT_TO_WORD(iN),8)+16#0009;
				EXIT;
			END_IF
			IrAngle_O3O4O6:=ACOS((lrLCirDis_pt3pt4*lrLCirDis_pt3pt4+lrLCirDis_pt4pt6*lrLCirDis_pt4pt6-lrLCirDis_pt3pt6*lrLCirDis_pt3pt6)/(2*lrLCirDis_pt3pt4*lrLCirDis_pt4pt6));
			IF ABS((lrLCirDis_pt3pt4*lrLCirDis_pt3pt4+lrLCirDis_pt4pt6*lrLCirDis_pt4pt6-lrLCirDis_pt3pt6*lrLCirDis_pt3pt6)/(2*lrLCirDis_pt3pt4*lrLCirDis_pt4pt6))>1 THEN
				wResult:=SHL(INT_TO_WORD(iN),8)+16#00010;
				EXIT;
			END_IF
			IrAngle_O2O4P:=ASIN((ABS(pstStMechanicalParam_03^.lrD2-pstStMechanicalParam_03^.lrD4))/(2*lrLCirDis_pt2pt4));
			IF ABS((ABS(pstStMechanicalParam_03^.lrD2-pstStMechanicalParam_03^.lrD4))/(2*lrLCirDis_pt2pt4))>1 THEN
				wResult:=SHL(INT_TO_WORD(iN),8)+16#00011;
				EXIT;
			END_IF
			IrAngle_O2O4O6:=ACOS((lrLCirDis_pt2pt4*lrLCirDis_pt2pt4+lrLCirDis_pt4pt6*lrLCirDis_pt4pt6-lrLCirDis_pt2pt6*lrLCirDis_pt2pt6)/(2*lrLCirDis_pt2pt4*lrLCirDis_pt4pt6));
			IF ABS((lrLCirDis_pt2pt4*lrLCirDis_pt2pt4+lrLCirDis_pt4pt6*lrLCirDis_pt4pt6-lrLCirDis_pt2pt6*lrLCirDis_pt2pt6)/(2*lrLCirDis_pt2pt4*lrLCirDis_pt4pt6))>1 THEN
				wResult:=SHL(INT_TO_WORD(iN),8)+16#00012;
				EXIT;
			END_IF
			IrAngle_NO4Q:=1.5*gc_lrPI-IrAngle_O6O4N-IrAngle_O2O4O6-IrAngle_O2O4P;(*圆4上需要计算的弧度*)
			IrAngle_ZO5W:=ATAN((pstStMechanicalParam_03^.lrY5-pstStMechanicalParam_03^.lrY3)/(pstStMechanicalParam_03^.lrX5-pstStMechanicalParam_03^.lrX3));
			IF pstStMechanicalParam_03^.lrx5=pstStMechanicalParam_03^.lrX3 THEN(*分母不能为零*)
				wResult:=SHL(INT_TO_WORD(iN),8)+16#00013;
				EXIT;
			END_IF
			IrAngle_WO5S:=gc_lrPI-IrAngle_ZO5W-IrAngle_HO3M;(*圆5上需要计算的弧度*)
			IrArc_UV:=IrAngle_UO2V*pstStMechanicalParam_03^.lrD2/2;(*圆2上需要计算的弧长*)
			IrArc_HI:=0.5*IrAngle_HO3I*pstStMechanicalParam_03^.lrD3;(*圆3上需要计算的弧长*)
			IrArc_NQ:=0.5*IrAngle_NO4Q*pstStMechanicalParam_03^.lrD4;(*圆4上需要计算的弧长*)
			IrArc_WS:=IrAngle_WO5S*(pstStMechanicalParam_03^.lrD5/2);(*圆5上需要进行的弧长*)
			IrIU:=SQRT(lrLCirDis_pt2pt3*lrLCirDis_pt2pt3-(((pstStMechanicalParam_03^.lrD2-pstStMechanicalParam_03^.lrD3)/2)*((pstStMechanicalParam_03^.lrD2-pstStMechanicalParam_03^.lrD3)/2)));
			IrQV:=SQRT(lrLCirDis_pt2pt4*lrLCirDis_pt2pt4-(((pstStMechanicalParam_03^.lrD2-pstStMechanicalParam_03^.lrD4)/2)*((pstStMechanicalParam_03^.lrD2-pstStMechanicalParam_03^.lrD4)/2)));
			IrHS:=((pstStMechanicalParam_03^.lrD3+pstStMechanicalParam_03^.lrD5)*IrHM)/pstStMechanicalParam_03^.lrD3;
			IrNT:=SQRT(lrLCirDis_pt4pt6*lrLCirDis_pt4pt6+(((pstStMechanicalParam_03^.lrD4-pstStMechanicalParam_03^.lrD6)/2)*((pstStMechanicalParam_03^.lrD4-pstStMechanicalParam_03^.lrD6)/2)));
			alrConstantLength[iN]:= IrArc_UV+IrArc_HI+IrArc_NQ+IrArc_WS+IrIU+IrQV+IrHS+IrNT;(*可变料长*)
			lrTotalLength:=alrConstantLength[iN]+i_pstStSysParam^.astStUnitParam_Save[iAxisId].lrPreReg_ConstVal;
			(*2024.7.11.164906+*)

			IF i_xFilpSwitch THEN(*翻转架开关打开了|就把翻料架的料长加进去@一般一台机器只有一个翻料架*)
				IF i_pstStSysParam^.astStGrpParam_Save[i_iGrpId].byTurnOverAxisId=0 THEN(*=0|那个轴有翻料架值就直接累加*)
					lrTotalLength:=lrTotalLength+i_pstStSysParam^.astStUnitParam_Save[iAxisId].uiTurnOverFilmLenth;
				ELSE
					IF i_pstStSysParam^.astStGrpParam_Save[i_iGrpId].byTurnOverAxisId=iAxisId THEN(*就是输入的轴id@累加该轴的翻料架长度*)
						lrTotalLength:=lrTotalLength+i_pstStSysParam^.astStUnitParam_Save[iAxisId].uiTurnOverFilmLenth;
					END_IF
				END_IF
			END_IF

			IF iN=1 THEN
				lrTotalLength:=0;
				i_pstStSysParam^.astStUnitParam_Save[iAxisId].lrPreReg_Length_V:=0;
				i_pstStSysParam^.astStUnitParam_Save[iAxisId].lrFilmLengthFromPrevUnit:=lrTotalLength;
			ELSE
				i_pstStSysParam^.astStUnitParam_Save[iAxisId].lrFilmLengthFromPrevUnit:=lrTotalLength;
				i_pstStSysParam^.astStUnitParam_Save[iAxisId].lrPreReg_Length_V:= KS_LREAL_MOD(lrTotalLength, i_pstStSysParam^.astStUnitParam_Save[iAxisId].rGirth_PrnRoller);(*当前色预套准计算的值*)
				i_pstStSysParam^.astStUnitParam_Save[iAxisId].lrPreReg_Length_V:=i_pstStSysParam^.astStUnitParam_Save[iAxisId].rGirth_PrnRoller-i_pstStSysParam^.astStUnitParam_Save[iAxisId].lrPreReg_Length_V
									+i_pstStSysParam^.astStUnitParam_Save[iAxisId].lrPreReg_Adjust+i_pstStSysParam^.astStUnitParam_Save[i_aiGrpAxisList[iN-1]].lrPreReg_Length_V;

				(* 2020.9.11.152457|防止输入的修正值绝对值超出1个版周 *)
				WHILE i_pstStSysParam^.astStUnitParam_Save[iAxisId].lrPreReg_Length_V<0 DO
					i_pstStSysParam^.astStUnitParam_Save[iAxisId].lrPreReg_Length_V:= i_pstStSysParam^.astStUnitParam_Save[iAxisId].lrPreReg_Length_V+i_pstStSysParam^.astStUnitParam_Save[iAxisId].rGirth_PrnRoller;
				END_WHILE
				WHILE i_pstStSysParam^.astStUnitParam_Save[iAxisId].lrPreReg_Length_V>i_pstStSysParam^.astStUnitParam_Save[iAxisId].rGirth_PrnRoller DO
					i_pstStSysParam^.astStUnitParam_Save[iAxisId].lrPreReg_Length_V:= i_pstStSysParam^.astStUnitParam_Save[iAxisId].lrPreReg_Length_V-i_pstStSysParam^.astStUnitParam_Save[iAxisId].rGirth_PrnRoller;
				END_WHILE

			END_IF
		END_FOR
	4:(*定料长*)
		FOR iN:=1 TO i_iGrpAxisNum_Pu BY 1 DO
			iAxisId:= i_aiGrpAxisList[iN];

			i_pstStSysParam^.astStUnitParam_Save[iAxisId].lrFilmLengthFromPrevUnit:=i_pstStSysParam^.astStUnitParam_Save[iAxisId].lrPreReg_ConstVal;(*2022.6.24.110711 定料长=机组料长|还存在定料长变化的可能-未处理~~*)
			IF iN=1 THEN
				i_pstStSysParam^.astStUnitParam_Save[iAxisId].lrPreReg_Length_V:=0;
				i_pstStSysParam^.astStUnitParam_Save[iAxisId].lrFilmLengthFromPrevUnit:=0;
			ELSE
				(*该值由界面提供，不该赋值|2020.9.8.174713|Liu.yt*)
				i_pstStSysParam^.astStUnitParam_Save[iAxisId].lrPreReg_Length_V:= KS_LREAL_MOD(i_pstStSysParam^.astStUnitParam_Save[iAxisId].lrFilmLengthFromPrevUnit, i_pstStSysParam^.astStUnitParam_Save[iAxisId].rGirth_PrnRoller);(*当前色预套准计算的值*)
				(*没有增加修正量|2022.6.24.110718*)
				i_pstStSysParam^.astStUnitParam_Save[iAxisId].lrPreReg_Length_V:=i_pstStSysParam^.astStUnitParam_Save[iAxisId].rGirth_PrnRoller-i_pstStSysParam^.astStUnitParam_Save[iAxisId].lrPreReg_Length_V
									+i_pstStSysParam^.astStUnitParam_Save[iAxisId].lrPreReg_Adjust+i_pstStSysParam^.astStUnitParam_Save[i_aiGrpAxisList[iN-1]].lrPreReg_Length_V;
				(* 2020.9.11.152457|防止输入的修正值绝对值超出1个版周 *)
				WHILE i_pstStSysParam^.astStUnitParam_Save[iAxisId].lrPreReg_Length_V<0 DO
					i_pstStSysParam^.astStUnitParam_Save[iAxisId].lrPreReg_Length_V:= i_pstStSysParam^.astStUnitParam_Save[iAxisId].lrPreReg_Length_V+i_pstStSysParam^.astStUnitParam_Save[iAxisId].rGirth_PrnRoller;
				END_WHILE
				WHILE i_pstStSysParam^.astStUnitParam_Save[iAxisId].lrPreReg_Length_V>i_pstStSysParam^.astStUnitParam_Save[iAxisId].rGirth_PrnRoller  DO
					i_pstStSysParam^.astStUnitParam_Save[iAxisId].lrPreReg_Length_V:= i_pstStSysParam^.astStUnitParam_Save[iAxisId].lrPreReg_Length_V-i_pstStSysParam^.astStUnitParam_Save[iAxisId].rGirth_PrnRoller;
				END_WHILE

			END_IF
		END_FOR

	(*2026.08.27.095631*)
	5: (*欧诺+力达直压式|2023.07.10.142323||2023.11.17.101158||2026.08.26 重构||[AI修改20260827]rD0改由本轴版周长推算+包角负值改报错*)
    pstStMechanicalParam_05 := ADR(i_pastStMechanicalParamBuf^[5].abyBuf);

    (* --- 1. 输入参数有效性检查（统一返回 16#FF01） --- *)
    IF pstStMechanicalParam_05^.rX1 < 0.1 OR pstStMechanicalParam_05^.rY1 < 0.1 OR
       pstStMechanicalParam_05^.rX2 < 0.1 OR pstStMechanicalParam_05^.rX3 < 0.1 OR
       pstStMechanicalParam_05^.rX4 < 0.1 OR pstStMechanicalParam_05^.rY4 < 0.1 OR
       pstStMechanicalParam_05^.rY0 < 0.1 OR pstStMechanicalParam_05^.rY2 < 0.1 OR(*[AI修改20260829]检查项rL2_3→rY2|前者转动态派生,不再作静态输入检查*)
       pstStMechanicalParam_05^.rD1 < 0.1 OR(*[AI修改20260827]移除rD0项|版辊直径不再作为静态输入*)
       pstStMechanicalParam_05^.rD2 < 0.1 OR pstStMechanicalParam_05^.rD3 < 0.1 OR
       pstStMechanicalParam_05^.rD4 < 0.1 THEN
        wResult := 16#FF01;  (* 全局参数无效 *)
        RETURN;
    END_IF

    FOR iN := 1 TO i_iGrpAxisNum_Pu BY 1 DO
        iAxisId := i_aiGrpAxisList[iN];
        rPlateR := i_pstStSysParam^.astStUnitParam_Save[iAxisId].rGirth_PrnRoller/gc_lrPi/2.0;(*[AI修改20260827]版辊半径=本轴版周长/π/2|替代原静态rD0/2,几何随轴变化*)
        rY3 := pstStMechanicalParam_05^.rY0 + rPlateR + pstStMechanicalParam_05^.rD3/2;(*[AI修改20260829]辊3(D3)辊心高=动态|Y0+版半径+D3半径,随版径浮动|同原版2023.11算法(原rY5项)*)
        rL2_3 := pstStMechanicalParam_05^.rY2 - rY3;(*[AI修改20260829]辊2-3垂直中心距=动态派生|修正:辊2高度rY2为固定安装尺寸,原静态字段rL2_3删除*)

        (* --- 2. 圆心距计算 --- *)
        rd1 := SQRT(EXPT(pstStMechanicalParam_05^.rX1 - pstStMechanicalParam_05^.rX2, 2) +
                    EXPT(pstStMechanicalParam_05^.rY1 - pstStMechanicalParam_05^.rY0 -
                         rPlateR - pstStMechanicalParam_05^.rD3/2 -
                         rL2_3, 2));
        rd2 := SQRT(EXPT(pstStMechanicalParam_05^.rX3 - pstStMechanicalParam_05^.rX2, 2) +
                    EXPT(rL2_3, 2));
        rd3 := SQRT(EXPT(pstStMechanicalParam_05^.rX4 - pstStMechanicalParam_05^.rX3, 2) +
                    EXPT(pstStMechanicalParam_05^.rY4 - pstStMechanicalParam_05^.rY0 -
                         rPlateR - pstStMechanicalParam_05^.rD3/2, 2));
        rd4 := SQRT(EXPT(pstStMechanicalParam_05^.rX3 - pstStMechanicalParam_05^.rX1, 2) +
                    EXPT(pstStMechanicalParam_05^.rY1 - pstStMechanicalParam_05^.rY0 -
                         rPlateR - pstStMechanicalParam_05^.rD3/2, 2));
        rd5 := SQRT(EXPT(pstStMechanicalParam_05^.rX4 - pstStMechanicalParam_05^.rX2, 2) +
                    EXPT(pstStMechanicalParam_05^.rY4 - pstStMechanicalParam_05^.rY0 -
                         rPlateR - pstStMechanicalParam_05^.rD3/2 -
                         rL2_3, 2));

        (* --- 3. 圆心距为零检查 --- *)
        IF rd1 = 0 OR rd2 = 0 OR rd3 = 0 OR rd4 = 0 OR rd5 = 0 THEN
            wResult := SHL(INT_TO_WORD(iN), 8) + 16#0001;  (* 圆心距为零 *)
            EXIT;
        END_IF

        (* --- 4. 切线长度计算（允许临界零切线） --- *)
        IF rd1 >= (pstStMechanicalParam_05^.rD1/2 + pstStMechanicalParam_05^.rD2/2) THEN
            rLength1 := SQRT(EXPT(rd1, 2) - EXPT(pstStMechanicalParam_05^.rD1/2 + pstStMechanicalParam_05^.rD2/2, 2));
        ELSE
            wResult := SHL(INT_TO_WORD(iN), 8) + 16#0002;  (* 外切条件不满足 *)
            EXIT;
        END_IF

        IF rd2 >= ABS(pstStMechanicalParam_05^.rD3/2 - pstStMechanicalParam_05^.rD2/2) THEN
            rLength2 := SQRT(EXPT(rd2, 2) - EXPT(pstStMechanicalParam_05^.rD3/2 - pstStMechanicalParam_05^.rD2/2, 2));
        ELSE
            wResult := SHL(INT_TO_WORD(iN), 8) + 16#0003;  (* 内切条件不满足（D2-D3） *)
            EXIT;
        END_IF

        IF rd3 >= ABS(pstStMechanicalParam_05^.rD3/2 - pstStMechanicalParam_05^.rD4/2) THEN
            rLength3 := SQRT(EXPT(rd3, 2) - EXPT(pstStMechanicalParam_05^.rD3/2 - pstStMechanicalParam_05^.rD4/2, 2));
        ELSE
            wResult := SHL(INT_TO_WORD(iN), 8) + 16#0004;  (* 内切条件不满足（D3-D4） *)
            EXIT;
        END_IF

        (* --- 5. 圆心到切点距离 --- *)
        rCenter_To_tangent1 := SQRT(EXPT(rLength1, 2) + EXPT(pstStMechanicalParam_05^.rD1/2, 2));
        rCenter_To_tangent2 := SQRT(EXPT(rLength2, 2) + EXPT(pstStMechanicalParam_05^.rD3/2, 2));
        rCenter_To_tangent3 := SQRT(EXPT(rLength2, 2) + EXPT(pstStMechanicalParam_05^.rD2/2, 2));
        rCenter_To_tangent4 := SQRT(EXPT(rLength3, 2) + EXPT(pstStMechanicalParam_05^.rD4/2, 2));

        (* --- 6. 角度与弧长计算（带余弦值域校验） --- *)
        lrTemp := (EXPT(rd1, 2) + EXPT(pstStMechanicalParam_05^.rD2/2, 2) - EXPT(rCenter_To_tangent1, 2)) /
                  (2 * rd1 * pstStMechanicalParam_05^.rD2/2);
        IF ABS(lrTemp) > 1.0 THEN
            wResult := SHL(INT_TO_WORD(iN), 8) + 16#0005;  (* 角度1余弦超限 *)
            EXIT;
        END_IF
        rArc1 := ACOS(lrTemp);
        rAngle1 := rArc1 * 180 / gc_lrPi;

        lrTemp := (EXPT(rd1, 2) + EXPT(rd2, 2) - EXPT(rd4, 2)) / (2 * rd1 * rd2);
        IF ABS(lrTemp) > 1.0 THEN
            wResult := SHL(INT_TO_WORD(iN), 8) + 16#0006;  (* 角度2余弦超限 *)
            EXIT;
        END_IF
        rArc2 := ACOS(lrTemp);
        rAngle2 := rArc2 * 180 / gc_lrPi;

        lrTemp := (EXPT(rd2, 2) + EXPT(pstStMechanicalParam_05^.rD2/2, 2) - EXPT(rCenter_To_tangent2, 2)) /
                  (2 * rd2 * pstStMechanicalParam_05^.rD2/2);
        IF ABS(lrTemp) > 1.0 THEN
            wResult := SHL(INT_TO_WORD(iN), 8) + 16#0007;  (* 角度3余弦超限 *)
            EXIT;
        END_IF
        rArc3 := ACOS(lrTemp);
        rAngle3 := rArc3 * 180 / gc_lrPi;

        rAngle4 := 360 - rAngle1 - rAngle2 - rAngle3;
        IF rAngle4 < 0 THEN(*[AI修改20260827]D2包角为负=几何参数不自洽|仿CASE1/2/3改报错,不再钳零*)
            wResult := SHL(INT_TO_WORD(iN), 8) + 16#000B;  (* D2包角为负 *)
            EXIT;
        END_IF
        rArcLen1 := (gc_lrPi * rAngle4 * pstStMechanicalParam_05^.rD2/2) / 180;

        lrTemp := (EXPT(rd2, 2) + EXPT(pstStMechanicalParam_05^.rD3/2, 2) - EXPT(rCenter_To_tangent3, 2)) /
                  (2 * rd2 * pstStMechanicalParam_05^.rD3/2);
        IF ABS(lrTemp) > 1.0 THEN
            wResult := SHL(INT_TO_WORD(iN), 8) + 16#0008;  (* 角度5余弦超限 *)
            EXIT;
        END_IF
        rArc5 := ACOS(lrTemp);
        rAngle5 := rArc5 * 180 / gc_lrPi;

        lrTemp := (EXPT(rd2, 2) + EXPT(rd3, 2) - EXPT(rd5, 2)) / (2 * rd2 * rd3);
        IF ABS(lrTemp) > 1.0 THEN
            wResult := SHL(INT_TO_WORD(iN), 8) + 16#0009;  (* 角度6余弦超限 *)
            EXIT;
        END_IF
        rArc6 := ACOS(lrTemp);
        rAngle6 := rArc6 * 180 / gc_lrPi;

        lrTemp := (EXPT(rd3, 2) + EXPT(pstStMechanicalParam_05^.rD3/2, 2) - EXPT(rCenter_To_tangent4, 2)) /
                  (2 * rd3 * pstStMechanicalParam_05^.rD3/2);
        IF ABS(lrTemp) > 1.0 THEN
            wResult := SHL(INT_TO_WORD(iN), 8) + 16#000A;  (* 角度7余弦超限 *)
            EXIT;
        END_IF
        rArc7 := ACOS(lrTemp);
        rAngle7 := rArc7 * 180 / gc_lrPi;

        rAngle8 := 360 - rAngle5 - rAngle6 - rAngle7;
        IF rAngle8 < 0 THEN(*[AI修改20260827]D3包角为负=几何参数不自洽|仿CASE1/2/3改报错,不再钳零*)
            wResult := SHL(INT_TO_WORD(iN), 8) + 16#000C;  (* D3包角为负 *)
            EXIT;
        END_IF
        rArcLen2 := (gc_lrPi * rAngle8 * pstStMechanicalParam_05^.rD3/2) / 180;

        (* --- 7. 累加可变料长 --- *)
        alrConstantLength[iN] := rLength1 + rArcLen1 + rLength2 + rArcLen2 + rLength3;
        lrTotalLength := alrConstantLength[iN] + i_pstStSysParam^.astStUnitParam_Save[iAxisId].lrPreReg_ConstVal;

        (* --- 8. 翻转架逻辑（与CASE 1完全一致） --- *)
        IF i_xFilpSwitch THEN
            IF i_pstStSysParam^.astStGrpParam_Save[i_iGrpId].byTurnOverAxisId = 0 THEN
                lrTotalLength := lrTotalLength + i_pstStSysParam^.astStUnitParam_Save[iAxisId].uiTurnOverFilmLenth;
            ELSE
                IF i_pstStSysParam^.astStGrpParam_Save[i_iGrpId].byTurnOverAxisId = iAxisId THEN
                    lrTotalLength := lrTotalLength + i_pstStSysParam^.astStUnitParam_Save[iAxisId].uiTurnOverFilmLenth;
                END_IF
            END_IF
        END_IF

        (* --- 9. 预套准值计算（与其它CASE完全一致） --- *)
        IF iN = 1 THEN
            lrTotalLength := 0;
            i_pstStSysParam^.astStUnitParam_Save[iAxisId].lrPreReg_Length_V := 0;
            i_pstStSysParam^.astStUnitParam_Save[iAxisId].lrFilmLengthFromPrevUnit := lrTotalLength;
        ELSE
            i_pstStSysParam^.astStUnitParam_Save[iAxisId].lrFilmLengthFromPrevUnit := lrTotalLength;
            i_pstStSysParam^.astStUnitParam_Save[iAxisId].lrPreReg_Length_V :=
                KS_LREAL_MOD(lrTotalLength, i_pstStSysParam^.astStUnitParam_Save[iAxisId].rGirth_PrnRoller);
            i_pstStSysParam^.astStUnitParam_Save[iAxisId].lrPreReg_Length_V :=
                (i_pstStSysParam^.astStUnitParam_Save[iAxisId].rGirth_PrnRoller -
                 i_pstStSysParam^.astStUnitParam_Save[iAxisId].lrPreReg_Length_V) +
                i_pstStSysParam^.astStUnitParam_Save[iAxisId].lrPreReg_Adjust +
                i_pstStSysParam^.astStUnitParam_Save[i_aiGrpAxisList[iN-1]].lrPreReg_Length_V;

            WHILE i_pstStSysParam^.astStUnitParam_Save[iAxisId].lrPreReg_Length_V < 0 DO
                i_pstStSysParam^.astStUnitParam_Save[iAxisId].lrPreReg_Length_V :=
                    i_pstStSysParam^.astStUnitParam_Save[iAxisId].lrPreReg_Length_V +
                    i_pstStSysParam^.astStUnitParam_Save[iAxisId].rGirth_PrnRoller;
            END_WHILE
            WHILE i_pstStSysParam^.astStUnitParam_Save[iAxisId].lrPreReg_Length_V >
                  i_pstStSysParam^.astStUnitParam_Save[iAxisId].rGirth_PrnRoller DO
                i_pstStSysParam^.astStUnitParam_Save[iAxisId].lrPreReg_Length_V :=
                    i_pstStSysParam^.astStUnitParam_Save[iAxisId].lrPreReg_Length_V -
                    i_pstStSysParam^.astStUnitParam_Save[iAxisId].rGirth_PrnRoller;
            END_WHILE
        END_IF
    END_FOR
	6:(*2024.12.03.104056//秦华履带式柔印//Hou.N*)
		iUnitValid := 0;
		lrTemp_Qinhua := 0;
		lrPreReg_Len_V := 0;
		FOR iN:=1 TO i_iGrpAxisNum_Pu BY 1 DO
			iAxisId:= iN;
			pstStUnitParam_Save:= ADR(i_pstStSysParam^.astStUnitParam_Save[iAxisId]);
			pstStUnitParam_UnSave:= ADR(i_pstStSysParam^.astStUnitParam_UnSave[iAxisId]);
			pstStUnitParam_Save^.lrFilmLengthFromPrevUnit:= pstStUnitParam_Save^.lrPreReg_ConstVal;
			IF pstStUnitParam_Save^.xLinkage THEN
				IF iN=1 THEN//首色
					lrTotalLength:= 0;
					pstStUnitParam_Save^.lrPreReg_Length_V:= 0;
					pstStUnitParam_Save^.lrFilmLengthFromPrevUnit:= 0;
				ELSE
					IF NOT xUnitValid THEN
						pstStUnitParam_Save^.lrFilmLengthFromPrevUnit := pstStUnitParam_Save^.lrFilmLengthFromPrevUnit + lrTemp_Qinhua;
						lrTemp_Qinhua := 0;
					END_IF
					pstStUnitParam_Save^.lrPreReg_Length_V:= KS_LREAL_MOD(pstStUnitParam_Save^.lrFilmLengthFromPrevUnit,pstStUnitParam_Save^.rGirth_PrnRoller);
					pstStUnitParam_Save^.lrPreReg_Length_V:= (pstStUnitParam_Save^.rGirth_PrnRoller-pstStUnitParam_Save^.lrPreReg_Length_V) + (* 版向走料方向单方向运动的是余数部分 *)
									pstStUnitParam_Save^.lrPreReg_Adjust + (* 输入的修正值 *)
									i_pstStSysParam^.astStUnitParam_Save[iAxisId-1].lrPreReg_Length_V; (* 前一色已经运动过的量|相当于更新变化后的基准位置 *)

													(* 2020.9.11.152457|防止输入的修正值绝对值超出1个版周 *)
					WHILE pstStUnitParam_Save^.lrPreReg_Length_V<0 DO
						pstStUnitParam_Save^.lrPreReg_Length_V:= pstStUnitParam_Save^.lrPreReg_Length_V+pstStUnitParam_Save^.rGirth_PrnRoller;
					END_WHILE
					WHILE pstStUnitParam_Save^.lrPreReg_Length_V>pstStUnitParam_Save^.rGirth_PrnRoller DO
						pstStUnitParam_Save^.lrPreReg_Length_V:= pstStUnitParam_Save^.lrPreReg_Length_V-pstStUnitParam_Save^.rGirth_PrnRoller;
					END_WHILE

				END_IF

				xUnitValid := TRUE;
			ELSE
				xUnitValid := FALSE;
				lrTemp_Qinhua := pstStUnitParam_Save^.lrPreReg_ConstVal + lrTemp_Qinhua;
				IF iAxisId > 1 THEN
					pstStUnitParam_Save^.lrPreReg_Length_V := i_pstStSysParam^.astStUnitParam_Save[iAxisId-1].lrPreReg_Length_V;
				ELSE
					pstStUnitParam_Save^.lrPreReg_Length_V := 0;
				END_IF
			END_IF
		END_FOR

	7: (*2026.01.15.84747//增加机组式-品字型//Hou.N*)
		FOR iN:=1 TO i_iGrpAxisNum_Pu BY 1 DO
			iAxisId:= iN;
			pstStUnitParam_Save:= ADR(i_pstStSysParam^.astStUnitParam_Save[iAxisId]);
			pstStUnitParam_UnSave:= ADR(i_pstStSysParam^.astStUnitParam_UnSave[iAxisId]);
			IF iN=1 THEN//首色
				lrTotalLength:= 0;
				pstStUnitParam_Save^.lrPreReg_Length_V:= 0;
				pstStUnitParam_Save^.lrFilmLengthFromPrevUnit:= 0;
			ELSE
				pstStUnitParam_Save^.lrFilmLengthFromPrevUnit:=  pstStUnitParam_Save^.lrPreReg_ConstVal;
// 				rPrRadius:=i_pstStSysParam^.astStGrpParam_Save[1].rGirth_PrnRoller/2/gc_lrPI;
// 				rBrRadius:=i_pstStSysParam^.astStGrpParam_Save[1].rGirth_BottomRoller/2/gc_lrPI;
// 				rHypotenuse:=rPrRadius+rBrRadius;
// 				alrAngle_Br[iAxisId]:=ACOS(ABS(g_arFix_RightEdge[iAxisId]/rHypotenuse));
// 				alrArc_length_Br[iAxisId]:=rBrRadius*alrAngle_Br[iAxisId];
//				pstStUnitParam_Save^.lrFilmLengthFromPrevUnit := pstStUnitParam_Save^.lrFilmLengthFromPrevUnit+alrArc_length_Br[iAxisId];

				pstStUnitParam_Save^.lrPreReg_Length_V:= KS_LREAL_MOD(pstStUnitParam_Save^.lrFilmLengthFromPrevUnit,pstStUnitParam_Save^.rGirth_PrnRoller);
				pstStUnitParam_Save^.lrPreReg_Length_V:= (pstStUnitParam_Save^.rGirth_PrnRoller-pstStUnitParam_Save^.lrPreReg_Length_V) + (* 版向走料方向单方向运动的是余数部分 *)
								pstStUnitParam_Save^.lrPreReg_Adjust + (* 输入的修正值 *)
								i_pstStSysParam^.astStUnitParam_Save[iAxisId-1].lrPreReg_Length_V; (* 前一色已经运动过的量|相当于更新变化后的基准位置 *)

												(* 2020.9.11.152457|防止输入的修正值绝对值超出1个版周 *)
				WHILE pstStUnitParam_Save^.lrPreReg_Length_V<0 DO
					pstStUnitParam_Save^.lrPreReg_Length_V:=pstStUnitParam_Save^.lrPreReg_Length_V+pstStUnitParam_Save^.rGirth_PrnRoller;
				END_WHILE
				WHILE pstStUnitParam_Save^.lrPreReg_Length_V>pstStUnitParam_Save^.rGirth_PrnRoller DO
					pstStUnitParam_Save^.lrPreReg_Length_V:= pstStUnitParam_Save^.lrPreReg_Length_V-pstStUnitParam_Save^.rGirth_PrnRoller;
				END_WHILE

			END_IF
		END_FOR
	ELSE;
	END_CASE
ELSE
	wResult:=16#FFFF;
END_IF

KS_CalcForPreRegister:= wResult;

(* ---- KS_GetAxisInitPhaseWhenPreRegister.st ---- *)
(*@CES
Name=KS_GetAxisInitPhaseWhenPreRegister
Type=FunctionBlock
TypeGuid=6f9dac99-8de1-4efc-8465-68ac443b7d08
Guid=f2256f17-a4f2-4244-aed7-c9a2efcbad83
HasDeclaration=True
HasImplementation=True
*)
{DECLARATION}
FUNCTION KS_GetAxisInitPhaseWhenPreRegister : BOOL
(*只处理了联动轴的*)
(*预套准时轴的初始相位初始位置处理方法|默认就是手动转动*)
VAR_INPUT
	i_byAxisInitPhaseTypeWhenPreRegister:BYTE;(*预套准时轴初始相位方式选择|默认手动转到mark线位置|=1 自动记忆初始相位解放双手*)
	i_xFlag_CanSaveData:BOOL;(*可以保存数据标志@只有再type=1时起作用*)
	(*一些按钮输入@需要外部清零作为沿触发*)
	i_xBtn_SaveAllData:BOOL;(*全部保存*)
	i_xBtn_SaveProtionData:BOOL;(*部分保存*)
	i_xBtn_SaveCancel:BOOL;(*取消按钮*)
	i_xBtn_DisHmi:BOOL;(*界面显示按钮*)
	(*轴的一些参数*)
	i_iGrpAxisNum_Pu: INT;(*色组轴的数量|*)
	i_aiGrpAxisList: ARRAY [1..MAX_UNIT_NUM] OF INT;(*系内所有轴的id列表,色组部分已经按照从小到大的顺序排序了，之后的是牵引|*)
	i_pstStSysParam: POINTER TO StSysParam;
//	i_pastStPTSts: POINTER TO ARRAY [1..MAX_UNIT_NUM] OF StPTSts;(*PT运动轴的状态|*)
	(*一些状态输出*)
	i_pxInitPhaseHmiSts:POINTER TO BOOL;(*初始相位操作界面状态标志位*)
	i_pxFlag_SaveAll:POINTER TO BOOL;(*全部保存标志*)
	i_pxFlag_SaveProtion:POINTER TO BOOL;(*部分保存标志*)
END_VAR
VAR
	iN: INT;
	iUnitId: INT;
//	pstStPTSts: POINTER TO StPTSts;(*PT运动轴的状态|*)
	xInitPhaseHmiSts: BOOL;
	xFlag_SaveAll: BOOL;
	xFlag_SaveProtion: BOOL;

	axInitPhaseValid:ARRAY [1..MAX_UNIT_NUM] OF BOOL;(*初始相位有效*)
	axNeedUpdate:ARRAY [1..MAX_UNIT_NUM] OF BOOL;(*需要更新的标志*)
	axUpdateDne:ARRAY [1..MAX_UNIT_NUM] OF BOOL;(*更新完成的标志*)
	axUpdateFailed:ARRAY [1..MAX_UNIT_NUM] OF BOOL;(*更新失败的标志*)
	xUpdateData: BOOL;(*更新数据标志*)
	xUpdateDne: BOOL;(*更新完成*)
	xFlag_CanSaveData: BOOL;(*可以保存数据*)
	xResetAxisFlag: BOOL;
END_VAR
{IMPLEMENTATION}
IF i_pxInitPhaseHmiSts<>0 THEN
	xInitPhaseHmiSts:=i_pxInitPhaseHmiSts^;
END_IF
IF i_pxFlag_SaveAll<>0 THEN
	xFlag_SaveAll:=i_pxFlag_SaveAll^;
END_IF
IF i_pxFlag_SaveProtion<>0 THEN
	xFlag_SaveProtion:=i_pxFlag_SaveProtion^;
END_IF

xFlag_CanSaveData:=i_xFlag_CanSaveData;

IF i_pstStSysParam<>0 THEN
	CASE i_byAxisInitPhaseTypeWhenPreRegister OF
		1:(*自动记忆初始相位解放双手*)

			(*获取状态位*)
			FOR iN:=1 TO i_iGrpAxisNum_Pu BY 1DO
				iUnitId:=i_aiGrpAxisList[iN];

				axInitPhaseValid[iUnitId]:=i_pstStSysParam^.astStUnitParam_Save[iUnitId].byPhaseState.0;
				axNeedUpdate[iUnitId]:=i_pstStSysParam^.astStUnitParam_Save[iUnitId].byPhaseState.1;
				axUpdateDne[iUnitId]:=i_pstStSysParam^.astStUnitParam_Save[iUnitId].byPhaseState.4;
				axUpdateFailed[iUnitId]:=i_pstStSysParam^.astStUnitParam_Save[iUnitId].byPhaseState.5;
			END_FOR

			(*按钮处理|*)
			IF NOT xFlag_SaveAll AND
				NOT xFlag_SaveProtion THEN(*存储标志无效的时候检测按钮输入*)
				(*全部更新按钮@保证互斥*)
				IF i_xBtn_SaveAllData THEN
					xFlag_SaveAll:=TRUE;
					xResetAxisFlag:=TRUE;(*复位轴标志@重新开始*)
				END_IF
				(*部分更新按钮@保证互斥*)
				IF NOT xFlag_SaveAll THEN
					IF i_xBtn_SaveProtionData THEN
						xFlag_SaveProtion:=TRUE;
						xResetAxisFlag:=TRUE;(*复位轴标志@重新开始*)
					END_IF
				END_IF
			END_IF

			(*界面显示按钮*)
			IF i_xBtn_DisHmi THEN
				xInitPhaseHmiSts:=TRUE;(*界面显示*)
			END_IF
			(*取消按钮*)
			IF i_xBtn_SaveCancel THEN
				xInitPhaseHmiSts:=FALSE;(*取消界面*)
			END_IF

			FOR iN:=1 TO i_iGrpAxisNum_Pu BY 1DO
				iUnitId:=i_aiGrpAxisList[iN];

				(*判断当前轴是否保存过初始版辊位置*)
				IF i_pstStSysParam^.astStUnitParam_Save[iUnitId].iPhase_InstallPlate<>0 THEN
					axInitPhaseValid[iUnitId]:=TRUE;
				ELSE
					axInitPhaseValid[iUnitId]:=FALSE;
				END_IF

				(*逻辑处理*)
				xUpdateData:=FALSE;
				IF xFlag_SaveAll THEN(*全部更新@2023.10.14.162459*)
					IF i_pstStSysParam^.astStUnitParam_Save[iUnitId].xLinkage THEN(*只要是联动的就更新*)
						xUpdateData:=TRUE;
						axNeedUpdate[iUnitId]:=TRUE;(*需要更新标志*)
					ELSE
						axNeedUpdate[iUnitId]:=FALSE;(*清除标志*)
					END_IF
				ELSIF xFlag_SaveProtion THEN(*部分更新@2023.10.14.162456*)
					IF i_pstStSysParam^.astStUnitParam_Save[iUnitId].xLinkage AND
						(NOT axInitPhaseValid[iUnitId]) THEN(*没有保存的进行更新*)
						xUpdateData:=TRUE;
						axNeedUpdate[iUnitId]:=TRUE;(*需要更新标志*)
					ELSE
						axNeedUpdate[iUnitId]:=FALSE;(*清除标志*)
					END_IF
				ELSE(*更新完了\不需要更新|清除一些标志*)
					axNeedUpdate[iUnitId]:=FALSE;(*清除标志*)
				END_IF

				IF NOT xInitPhaseHmiSts OR (*界面关闭的时候清除标志位*)
					xResetAxisFlag THEN(*重新开始*)
					axUpdateDne[iUnitId]:=FALSE;(*更新成功标志清除*)
					axUpdateFailed[iUnitId]:=FALSE;(*更新失败标志清除*)
				END_IF

				IF axUpdateDne[iUnitId] OR(*更新成功|都不再更新*)
					axUpdateFailed[iUnitId] THEN(*更新失败|都不再更新*)
					xUpdateData:=FALSE;
				END_IF

				(*需要更新位置*)
				IF xUpdateData THEN
					IF xFlag_CanSaveData THEN(*可以保存数据*)
						i_pstStSysParam^.astStUnitParam_Save[iUnitId].iPhase_InstallPlate:=
								KS_GetPhaseValue(i_pstStSysParam^.astStUnitParam_UnSave[iUnitId].wVirTual_Cnt,gc_iVirEncPPR);
						IF i_pstStSysParam^.astStUnitParam_Save[iUnitId].iPhase_InstallPlate=0 THEN(*保证保存的值非零*)
							i_pstStSysParam^.astStUnitParam_Save[iUnitId].iPhase_InstallPlate:=1;
						END_IF
						(*非法值判断*)
						IF i_pstStSysParam^.astStUnitParam_Save[iUnitId].iPhase_InstallPlate>0 AND
							i_pstStSysParam^.astStUnitParam_Save[iUnitId].iPhase_InstallPlate<gc_iVirEncPPR THEN(*值合法*)
							axUpdateDne[iUnitId]:=TRUE;(*更新完成*)
						ELSE
							axUpdateFailed[iUnitId]:=TRUE;(*更新失败*)
						END_IF
					ELSE(*不能保存数据|置位失败标志*)
						axUpdateFailed[iUnitId]:=TRUE;(*更新失败*)
					END_IF
				END_IF

			END_FOR

			(*处理整机标志位*)
			FOR iN:=1 TO i_iGrpAxisNum_Pu BY 1DO
				iUnitId:=i_aiGrpAxisList[iN];

				xUpdateDne:=(axUpdateDne[iUnitId] OR axUpdateFailed[iUnitId]);
				IF xFlag_SaveAll OR(*全部更新*)
					xFlag_SaveProtion(*部分更新*)THEN
					IF axNeedUpdate[iUnitId] THEN
						IF xUpdateDne THEN(*更新完成了*);
						ELSE
							EXIT;
						END_IF
					END_IF

					IF iN=i_iGrpAxisNum_Pu THEN(*能走到这里说明都完成了*)
						xFlag_SaveAll:=FALSE;
						xFlag_SaveProtion:=FALSE;
					END_IF
				END_IF
			END_FOR

			(*输出状态位*)
			FOR iN:=1 TO i_iGrpAxisNum_Pu BY 1DO
				iUnitId:=i_aiGrpAxisList[iN];
				i_pstStSysParam^.astStUnitParam_Save[iUnitId].byPhaseState.0:=axInitPhaseValid[iUnitId];
				i_pstStSysParam^.astStUnitParam_Save[iUnitId].byPhaseState.1:=axNeedUpdate[iUnitId];
				i_pstStSysParam^.astStUnitParam_Save[iUnitId].byPhaseState.4:=axUpdateDne[iUnitId];
				i_pstStSysParam^.astStUnitParam_Save[iUnitId].byPhaseState.5:=axUpdateFailed[iUnitId];
				(*清除无效位*)
				i_pstStSysParam^.astStUnitParam_Save[iUnitId].byPhaseState.2:=FALSE;
				i_pstStSysParam^.astStUnitParam_Save[iUnitId].byPhaseState.3:=FALSE;
				i_pstStSysParam^.astStUnitParam_Save[iUnitId].byPhaseState.6:=FALSE;
				i_pstStSysParam^.astStUnitParam_Save[iUnitId].byPhaseState.7:=FALSE;
			END_FOR

			IF NOT xInitPhaseHmiSts THEN(*界面关闭的时候清除标志位*)
				xFlag_SaveAll:=FALSE;
				xFlag_SaveProtion:=FALSE;
			END_IF
	ELSE(*默认方案*)
		FOR iN:=1 TO i_iGrpAxisNum_Pu BY 1DO
			iUnitId:=i_aiGrpAxisList[iN];

(*这里就不清零@2025.1.12.175804
KS_ReloadPreRegValue 这里加了大条件*)
(*			pstStAxisParam^.iPhase_InstallPlate:=0;(*清零这个值*)*)
			(*一些参数清除*)
			i_pstStSysParam^.astStUnitParam_Save[iUnitId].byPhaseState:=0;
		END_FOR
		xInitPhaseHmiSts:=FALSE;(*取消界面*)
		xFlag_SaveAll:=FALSE;(*全部保存标志*)
		xFlag_SaveProtion:=FALSE;(*部分保存标志*)
	END_CASE
END_IF

(*状态输出*)
IF i_pxInitPhaseHmiSts<>0 THEN
	i_pxInitPhaseHmiSts^:=xInitPhaseHmiSts;
END_IF
IF i_pxFlag_SaveAll<>0 THEN
	i_pxFlag_SaveAll^:=xFlag_SaveAll;
END_IF
IF i_pxFlag_SaveProtion<>0 THEN
	i_pxFlag_SaveProtion^:=xFlag_SaveProtion;
END_IF

(* ---- KS_GetCorrect_PreRegister_Auto.st ---- *)
(*@CES
Name=KS_GetCorrect_PreRegister_Auto
Type=FunctionBlock
TypeGuid=6f9dac99-8de1-4efc-8465-68ac443b7d08
Guid=3dff30e1-2ce5-4884-8d32-0e4848e202b7
HasDeclaration=True
HasImplementation=True
*)
{DECLARATION}
FUNCTION KS_GetCorrect_PreRegister_Auto : BOOL(*自动获取预套准修正量|
											    根据套色调整量获得*)
VAR_INPUT
	i_xAutoGetCorr:BOOL;(*自动获取预套准修正量标志|做完预套准后第一次印刷执行*)
	i_pxWrPreRegisterCorr:POINTER TO BOOL;(*写入到预套准修正值中标志*)
	i_iGrpAxisNum_Pu: INT; (*色组轴数量*)
	i_paiGrpAxisList: POINTER TO ARRAY [1..MAX_UNIT_NUM] OF INT; (*系内所有轴的列表*)
	i_pstStSysParam: POINTER TO StSysParam;
	i_iGrpId:int;(*系号*)
	i_palrTotalCorrectVal:POINTER TO ARRAY [1..MAX_UNIT_NUM] OF LREAL;(*总的修正量|mm*)
	i_palrTotalAdjustVal_V:POINTER TO ARRAY [1..MAX_UNIT_NUM] OF LREAL;(*套色总的调整量|mm*)
END_VAR
VAR
	iN:INT;
	iAxisId:INT;
	lrTotalAdjustVal: LREAL;(*总的调整量|单位都是um*)
	lrTotalAdjustValLastAxis: LREAL;(*上个轴的调整量*)
END_VAR
{IMPLEMENTATION}
IF i_paiGrpAxisList<>0 AND
	i_pstStSysParam<>0 AND
	i_palrTotalCorrectVal<>0 AND
	i_pxWrPreRegisterCorr<>0 AND
	i_palrTotalAdjustVal_V<>0 THEN
	IF i_pstStSysParam^.astStGrpParam_UnSave[i_iGrpId].xFlag_Print AND (*印刷时候我们才进行统计*)
		i_xAutoGetCorr THEN
		FOR iN:=1 TO MAX_UNIT_NUM BY 1 DO
			i_palrTotalCorrectVal^[iN]:=0;
		END_FOR

		lrTotalAdjustValLastAxis:=0;
		FOR iN:=1 TO i_iGrpAxisNum_Pu BY 1 DO
			iAxisId:=i_paiGrpAxisList^[iN];
		(*将以下部分总和起来就应该是总的调整量*)
			IF i_pstStSysParam^.astStUnitParam_Save[iAxisId].xLinkage THEN(*只统计联动轴*)
				lrTotalAdjustVal:=i_palrTotalAdjustVal_V^[iAxisId]-lrTotalAdjustValLastAxis;
				(*2021.6.16.084129 记录上个轴的调整量|计算需要的修正量*)
				lrTotalAdjustValLastAxis:=i_palrTotalAdjustVal_V^[iAxisId];
				i_palrTotalCorrectVal^[iAxisId]:=lrTotalAdjustVal/1000;
			END_IF
		END_FOR
	END_IF

	(*写入到预套准修正量中*)
	IF i_pxWrPreRegisterCorr^ THEN
		FOR iN:=1 TO i_iGrpAxisNum_Pu BY 1 DO
			iAxisId:=i_paiGrpAxisList^[iN];
			i_pstStSysParam^.astStUnitParam_Save[iAxisId].lrPreReg_Adjust:=i_pstStSysParam^.astStUnitParam_Save[iAxisId].lrPreReg_Adjust+
												i_palrTotalCorrectVal^[iAxisId];
		END_FOR
	END_IF
	i_pxWrPreRegisterCorr^:=FALSE;
END_IF

(* ---- KS_GetPhaseValue.st ---- *)
(*@CES
Name=KS_GetPhaseValue
Type=FunctionBlock
TypeGuid=6f9dac99-8de1-4efc-8465-68ac443b7d08
Guid=4208271a-275a-4ef9-bf83-b8f9c218fcae
HasDeclaration=True
HasImplementation=True
*)
{DECLARATION}
FUNCTION KS_GetPhaseValue : INT(*获取相位值@0--7999变化*)
VAR_INPUT
	i_wVirtualCnt:WORD;(*获取的虚拟码盘值0--65535变化*)
	i_iVirEncPPR:INT;(*一圈的脉冲数*)
END_VAR
VAR
	iVirtualCnt: INT;
	iVirtualPan_1Cycle:INT:=8000;
END_VAR
{IMPLEMENTATION}
iVirtualCnt:=WORD_TO_INT(i_wvirtualCnt);
iVirtualPan_1Cycle:=i_iVirEncPPR;
IF iVirtualPan_1Cycle=0 THEN
	iVirtualPan_1Cycle:=8000;
END_IF
IF iVirtualCnt>=0 AND
	iVirtualCnt<=iVirtualPan_1Cycle-1 THEN;
ELSE
	IF iVirtualCnt<0 THEN(*小于0*)
		REPEAT
			iVirtualCnt:=iVirtualCnt+iVirtualPan_1Cycle;
		UNTIL
			iVirtualCnt>=0
		END_REPEAT
	ELSE(*大于0*)
		iVirtualCnt:=iVirtualCnt MOD iVirtualPan_1Cycle;
	END_IF
END_IF
KS_GetPhaseValue:=iVirtualCnt;

(* ---- KS_JudgeMotorSts.st ---- *)
(*@CES
Name=KS_JudgeMotorSts
Type=FunctionBlock
TypeGuid=6f9dac99-8de1-4efc-8465-68ac443b7d08
Guid=a5e3ced4-c2da-4f83-ae84-e1a255808c54
HasDeclaration=True
HasImplementation=True
*)
{DECLARATION}
FUNCTION KS_JudgeMotorSts : BYTE(*判断电机状态函数|0 停止 1 运动*)
(*检测10个周期规划速度在一定阈值内则认为处于停止状态|*)
VAR_INPUT
	i_rMotorVel_FeedBack:REAL;(*反馈电机速度|PTsts反馈*)
	i_iThreshold:INT;(*判断的阈值|单位好像是脉冲*)
	i_iCycleNum_InStop:INT;(*处于停止的周期次数|这么多周期都处于阈值内就认为是停止了*)
	i_piCycleCnt_Stop:POINTER TO INT;(*处于停止阈值的周期计数*)
END_VAR
VAR
	iCycleCnt_Stop: INT;
	byMotorSts:BYTE;
END_VAR

{IMPLEMENTATION}
IF i_piCycleCnt_Stop<>0 THEN
	iCycleCnt_Stop:=i_piCycleCnt_Stop^;
END_IF

IF ABS(i_rMotorVel_FeedBack)<i_iThreshold THEN
	IF iCycleCnt_Stop<i_iCycleNum_InStop THEN
		iCycleCnt_Stop:=iCycleCnt_Stop+1;
	END_IF
ELSE
	iCycleCnt_Stop:=0;
END_IF

IF iCycleCnt_Stop>=i_iCycleNum_InStop THEN(*超过周期设定值|*)
	byMotorSts:=0;
ELSE
	byMotorSts:=1;
END_IF

IF i_piCycleCnt_Stop<>0 THEN
	i_piCycleCnt_Stop^:=iCycleCnt_Stop;
END_IF

KS_JudgeMotorSts:=byMotorSts;

(* ---- KS_LREAL_MOD.st ---- *)
(*@CES
Name=KS_LREAL_MOD
Type=FunctionBlock
TypeGuid=6f9dac99-8de1-4efc-8465-68ac443b7d08
Guid=d022a916-afa9-4b10-a8f8-a759c4e31692
HasDeclaration=True
HasImplementation=True
*)
{DECLARATION}
FUNCTION KS_LREAL_MOD : LREAL
VAR_INPUT
	i_lrData		: LREAL; (* 被模数 *)
	i_lrDividedBy	: LREAL; (* 模数 *)
END_VAR
VAR
	lrResult		: LREAL;
	diQuotient		: DINT; (* 整数的商/可能存在四舍五入 *)
	lrTmpValue		: LREAL;
END_VAR

{IMPLEMENTATION}
lrResult:= 0;
IF i_lrDividedBy<>0 AND i_lrData<>0 THEN
	diQuotient:= LREAL_TO_DINT(i_lrData/i_lrDividedBy); (* 由于LREAL_TO_DINT()会四舍五入,所以反算回去记得要考虑两边值 *)
	lrTmpValue:= i_lrDividedBy*diQuotient; (* 反算回去的结果 *)
	IF (i_lrData>0 AND lrTmpValue>i_lrData) OR
		(i_lrData<0 AND lrTmpValue<i_lrData) THEN
		(* 说明diQuotient被四舍五入了/比正值大/比负值小 *)
		IF diQuotient>0 THEN
			diQuotient:= diQuotient-1;
		ELSE
			diQuotient:= diQuotient+1;
		END_IF
	END_IF
	lrResult:= i_lrData-i_lrDividedBy*diQuotient;
END_IF
KS_LREAL_MOD:= lrResult;

(* ---- KS_ReloadPreRegValue.st ---- *)
(*@CES
Name=KS_ReloadPreRegValue
Type=FunctionBlock
TypeGuid=6f9dac99-8de1-4efc-8465-68ac443b7d08
Guid=57fb531d-4a0f-4c52-9839-1f16e0b31222
HasDeclaration=True
HasImplementation=True
*)
{DECLARATION}
FUNCTION KS_ReloadPreRegValue : INT
(*2022.9.8.120612 只计算联动轴*)
(*2023.6.25.151146 计算的时候取消了联动条件*)
(*2023.10.16.171750 重新启用aiVirEnc_AlignMarkToSamePosition变量作为自动对其mark线位置*)
(*2025.1.14.081723 单色预套功能还要再减去当前色的预套准量*)
(*2025.1.15.125933 1色也会计算调整量*)
VAR_INPUT
	i_iGrpId: INT;
	i_iGrpAxisNum_Pu: INT;
	i_aiGrpAxisList: ARRAY [1..MAX_UNIT_NUM] OF INT;
	i_pstStSysParam: POINTER TO StSysParam;
	i_pawAxisVirtualCnt: POINTER TO ARRAY [1..MAX_UNIT_NUM] OF WORD; (* 2021.6.25.104504/增加的虚拟编码器原始值输入 *)
	i_pawAxisVirtualSts: POINTER TO ARRAY [1..MAX_UNIT_NUM] OF WORD; (* 2021.6.25.104504/增加的虚拟编码器原始值输入 *)
	i_palrMovementResult: POINTER TO ARRAY [1..MAX_UNIT_NUM] OF LREAL;
	i_piDeltaPhase_MarkPos_FirstLinkage:POINTER TO INT;(*监控使用-第一个非手动预套的轴的信息@2025.1.12.183900*)
END_VAR
VAR
	iN: INT;
	iUnitId: INT;
	pstStAxisParam_FirstValidAxis: POINTER TO StUnitParam_Save;

//	pstStPTSts_FirstValidAxis: POINTER TO StPTSts;
//	pstStPTSts: POINTER TO StPTSts;

	iLastServoOnAxisId: INT;
	iFirstValidAxisId: INT;

	aiVirEnc_AxisResult: ARRAY [1..MAX_UNIT_NUM] OF INT;
	aiVirEnc_PlatePositionOffset: ARRAY [1..MAX_UNIT_NUM] OF INT; (*装版位置绝对差*)
	aiVirEnc_AlignMarkToSamePosition: ARRAY [1..MAX_UNIT_NUM] OF INT; (*对齐码刻线要移动的脉冲数*)
	aiVirEnc_AxisPreRegister: ARRAY [1..MAX_UNIT_NUM] OF INT;

	(*2025.1.12.180103*)
	iDeltaPhase_MarkPos_NotManuPreRegister1st:INT:=0;(*第一个不是手动预套的轴 距离mark位置的相位值@初值给个特殊值*)
END_VAR
{IMPLEMENTATION}
IF (i_iGrpId=1 OR i_iGrpId=2) AND
	(i_iGrpAxisNum_Pu>=1 AND i_iGrpAxisNum_Pu<=MAX_UNIT_NUM) AND
	i_pstStSysParam<>0 AND
	i_palrMovementResult<>0 THEN
	;
	FOR iN:=1 TO MAX_UNIT_NUM BY 1 DO
		aiVirEnc_PlatePositionOffset[iN]:= 0;
		aiVirEnc_AlignMarkToSamePosition[iN]:= 0;
		aiVirEnc_AxisPreRegister[iN]:= 0;
		aiVirEnc_AxisResult[iN]:= 0;
		i_palrMovementResult^[iN]:= 0;
	END_FOR

	(*2025.1.15.132938 移动*)
	(*先计算第一个非手动预套的轴联动色,当前位置距离mark线的值*)
	(*iPhase_InstallPlate 变量作为记录预套前的mark位置,用于实现单轴的预套准*)
	iDeltaPhase_MarkPos_NotManuPreRegister1st:=gc_iVirEncPPR;(*初值给个特殊值*)
	IF i_pstStSysParam^.astStGrpParam_Save[i_iGrpId].xPreRegisterAxisId_Manu THEN(*2025.1.14.142427 单轴预套的时候*)
		IF iDeltaPhase_MarkPos_NotManuPreRegister1st = gc_iVirEncPPR THEN(*第一个非手动预套的轴标记记录*)
			FOR iN:=1 TO i_iGrpAxisNum_Pu BY 1 DO
				iUnitId:= i_aiGrpAxisList[iN];

//				pstStPTSts:= ADR(i_pastStPTSts^[iAxisId]);
				(*预套准本身要走的量@后面计算要用*)

				aiVirEnc_AxisPreRegister[iUnitId]:=
					LREAL_TO_INT(i_pstStSysParam^.astStUnitParam_Save[iUnitId].lrPreReg_Length_V/ i_pstStSysParam^.astStUnitParam_Save[iUnitId].rGirth_PrnRoller * gc_iVirEncPPR);
				IF NOT i_pstStSysParam^.astStUnitParam_Save[iUnitId].xPreRegisterValid_Manu THEN
					iDeltaPhase_MarkPos_NotManuPreRegister1st:=(*当前位置-记录的mark位置*)
						KS_GetPhaseValue(i_pawAxisVirtualCnt^[iUnitId],gc_iVirEncPPR)-i_pstStSysParam^.astStUnitParam_Save[iUnitId].iPhase_InstallPlate;
					(*2025.1.14.081723 还要再减去当前色的预套准量*)
					iDeltaPhase_MarkPos_NotManuPreRegister1st:=iDeltaPhase_MarkPos_NotManuPreRegister1st-aiVirEnc_AxisPreRegister[iUnitId];

					IF iDeltaPhase_MarkPos_NotManuPreRegister1st<0 THEN
						iDeltaPhase_MarkPos_NotManuPreRegister1st:=iDeltaPhase_MarkPos_NotManuPreRegister1st+gc_iVirEncPPR;
					END_IF
					EXIT;
				END_IF
			END_FOR
		END_IF
	END_IF

	iFirstValidAxisId:= -1;
	iLastServoOnAxisId:= -1;
	FOR iN:=1 TO i_iGrpAxisNum_Pu BY 1 DO
		iUnitId:= i_aiGrpAxisList[iN];

//		pstStPTSts:= ADR(i_pastStPTSts^[iAxisId]);

			IF NOT (iFirstValidAxisId>=1 AND iFirstValidAxisId<=MAX_UNIT_NUM) THEN
				iFirstValidAxisId:= iUnitId;
			END_IF

			(*第一个轴不运动 从第二个轴开始运动*)
			IF iFirstValidAxisId>=1 AND iFirstValidAxisId<=MAX_UNIT_NUM THEN
				;
				pstStAxisParam_FirstValidAxis:= ADR(i_pstStSysParam^.astStUnitParam_Save[iFirstValidAxisId]);
//				pstStPTSts_FirstValidAxis:= ADR(i_pastStPTSts^[iFirstValidAxisId]);

				(*这个差值就是码刻线在同一位置，虚拟码盘的绝对差@未使用*)
				aiVirEnc_PlatePositionOffset[iUnitId]:=
					i_pstStSysParam^.astStUnitParam_Save[iUnitId].iPhase_InstallPlate-pstStAxisParam_FirstValidAxis^.iPhase_InstallPlate; (*和不动的第1色版装版位置绝对差*)

				(*预套准本身要走的量*)
				aiVirEnc_AxisPreRegister[iUnitId]:=
					LREAL_TO_INT(i_pstStSysParam^.astStUnitParam_Save[iUnitId].lrPreReg_Length_V/ i_pstStSysParam^.astStUnitParam_Save[iUnitId].rGirth_PrnRoller * gc_iVirEncPPR);

				(*2023.10.16.154812*)
				(*将码刻线对齐需要移动的脉冲数*)
				(*2025.1.12.171650 增加开关条件*)
				(*KS_FB_ProcPhaseOptReq 中增加逻辑实现预套时的mark位置记录*)
				IF i_pstStSysParam^.astStGrpParam_Save[i_iGrpId].byAxisInitPhaseTypeWhenPreRegister=1 THEN(*mark线和键槽固定相位时*)
					IF i_pstStSysParam^.astStUnitParam_Save[iUnitId].iPhase_InstallPlate<>0 AND(*有初始相位|计算需要执行的码盘数*)
						i_pawAxisVirtualSts^[iUnitId].12 THEN(*虚拟马盘是有效的*)
						aiVirEnc_AlignMarkToSamePosition[iUnitId]:=
							i_pstStSysParam^.astStUnitParam_Save[iUnitId].iPhase_InstallPlate-
							KS_GetPhaseValue(i_pawAxisVirtualCnt^[iUnitId],gc_iVirEncPPR);(*当前轴的位置偏差*)

						IF pstStAxisParam_FirstValidAxis^.iPhase_InstallPlate<>0 AND(*第一个轴有初始相位*)
							i_pawAxisVirtualSts^[iFirstValidAxisId].12 THEN(*虚拟马盘是有效的*)
							aiVirEnc_AlignMarkToSamePosition[iUnitId]:=
								aiVirEnc_AlignMarkToSamePosition[iUnitId]+
								KS_GetPhaseValue(i_pawAxisVirtualCnt^[iFirstValidAxisId],gc_iVirEncPPR)-
								pstStAxisParam_FirstValidAxis^.iPhase_InstallPlate;(*需要弥补的第一个轴位置偏差*)
						ELSE(*否则就舍弃掉*);
						END_IF
					ELSE
						aiVirEnc_AlignMarkToSamePosition[iUnitId]:=0;
					END_IF
				ELSE(*功能没开，这个计算值就写0*)
					(*iPhase_InstallPlate 变量作为记录预套前的mark位置,用于实现单轴的预套准*)
					(*先计算第一个非手动预套的轴联动色,当前位置距离mark线的值*)
					IF i_pstStSysParam^.astStUnitParam_Save[iUnitId].xPreRegisterValid_Manu THEN(*2025.1.14.142427 单轴预套的时候*)
						(*算出偏差*)
						IF iDeltaPhase_MarkPos_NotManuPreRegister1st<>gc_iVirEncPPR THEN
							aiVirEnc_AlignMarkToSamePosition[iUnitId]:=iDeltaPhase_MarkPos_NotManuPreRegister1st;
						END_IF
					ELSE
						aiVirEnc_AlignMarkToSamePosition[iUnitId]:=0;
					END_IF
				END_IF

				(*当前轴本身共走的量*)
				aiVirEnc_AxisResult[iUnitId]:=
					aiVirEnc_AlignMarkToSamePosition[iUnitId] +(*将对齐马克线的相位差加入到当前轴走的量里面|2023.10.16.171901*)
					aiVirEnc_AxisPreRegister[iUnitId] (*+
					aiVirEnc_AxisPreRegister[iLastServoOnAxisId]*); (* 2020.9.11.154445|取消掉之前的色组重复走了的值 *)

				WHILE aiVirEnc_AxisResult[iUnitId]<0 DO
					aiVirEnc_AxisResult[iUnitId]:= aiVirEnc_AxisResult[iUnitId]+gc_iVirEncPPR;
				END_WHILE
				WHILE aiVirEnc_AxisResult[iUnitId]>=gc_iVirEncPPR DO
					aiVirEnc_AxisResult[iUnitId]:= aiVirEnc_AxisResult[iUnitId]-gc_iVirEncPPR;
				END_WHILE

				(*将伺服电机需要走的量输出*)
				//2026.1.6.134228 | + | 不同机器类型处理
				IF g_iMachineryType	= MACHINERYTYPE_FELXO_INLINE_ONEBOTOMROLLER THEN
					i_palrMovementResult^[iUnitId]:=
							INT_TO_LREAL(aiVirEnc_AxisResult[iUnitId]) / INT_TO_LREAL(gc_iVirEncPPR) * i_pstStSysParam^.astStUnitParam_Save[iUnitId].rGirth_PrnRoller *
							(GC_LRMOTORPPR) * UINT_TO_LREAL(i_pstStSysParam^.astStUnitParam_Save[iUnitId].uiNum_BottomRoller) / UINT_TO_LREAL(i_pstStSysParam^.astStUnitParam_Save[iUnitId].uiDen_BottomRoller)/
							i_pstStSysParam^.astStUnitParam_Save[iUnitId].rGirth_BottomRoller;

					(*2020.9.8.155451 如果电机反转|我们需要将预套准输出值写反|Liu.yt*)
					IF i_pstStSysParam^.astStUnitParam_UnSave[iUnitId].xMotRev_BottomRoller THEN
						i_palrMovementResult^[iUnitId]:=
								-i_palrMovementResult^[iUnitId];
					END_IF
				ELSE
					i_palrMovementResult^[iUnitId]:=
							INT_TO_LREAL(aiVirEnc_AxisResult[iUnitId]) / INT_TO_LREAL(gc_iVirEncPPR) *
							(GC_LRMOTORPPR) * UINT_TO_LREAL(i_pstStSysParam^.astStUnitParam_Save[iUnitId].uiNum_PrnRoller) / UINT_TO_LREAL(i_pstStSysParam^.astStUnitParam_Save[iUnitId].uiDen_PrnRoller);

					(*2020.9.8.155451 如果电机反转|我们需要将预套准输出值写反|Liu.yt*)
					IF i_pstStSysParam^.astStUnitParam_UnSave[iUnitId].xMotRev_PrnRoller THEN
						i_palrMovementResult^[iUnitId]:=
								-i_palrMovementResult^[iUnitId];
					END_IF
				END_IF

			ELSE
				aiVirEnc_PlatePositionOffset[iUnitId]:= 0;
				aiVirEnc_AlignMarkToSamePosition[iUnitId]:= 0;
				aiVirEnc_AxisPreRegister[iUnitId]:= 0;
				aiVirEnc_AxisResult[iUnitId]:= 0;

				i_palrMovementResult^[iUnitId]:= 0;
			END_IF
			iLastServoOnAxisId:= iUnitId;

			IF NOT (iFirstValidAxisId>=1 AND iFirstValidAxisId<=MAX_UNIT_NUM) THEN
				iFirstValidAxisId:= iLastServoOnAxisId;
			END_IF
(*2023.6.25.151119屏蔽*)
(*		END_IF*)
	END_FOR
END_IF

(*2025.1.12.183940 增加一个监控*)
IF i_piDeltaPhase_MarkPos_FirstLinkage<>0 THEN
	IF iDeltaPhase_MarkPos_NotManuPreRegister1st<>gc_iVirEncPPR THEN
		i_piDeltaPhase_MarkPos_FirstLinkage^:=iDeltaPhase_MarkPos_NotManuPreRegister1st;
	END_IF
END_IF

(* ---- KS_SetMotionPovmd.st ---- *)
(*@CES
Name=KS_SetMotionPovmd
Type=FunctionBlock
TypeGuid=6f9dac99-8de1-4efc-8465-68ac443b7d08
Guid=ddeda59d-b720-4e82-aa52-b27576ad532a
HasDeclaration=True
HasImplementation=True
*)
{DECLARATION}
FUNCTION KS_SetMotionPovmd : INT(*2022.7.8.175801  新增加了PT模式使能切换模式
需要再pt功能初始化完成后有效即：设置pt模式和模态后使用*)
VAR_INPUT
	i_iStationId:INT;(*站号|*)
	i_xSetMotionPovmdEn:BOOL;(*设置PT使能模式使能*)
	i_wMotorEnMode:WORD;
	(*电机使能模式|0: 不使能 1: 使能 3: 使能后轴可以手动转动 4: 取消模式3状态
	3、4以为的值都不允许set
	实际应用下会3、4状态下切换*)
END_VAR
VAR
	iRtn:INT;
	wMode: WORD;
END_VAR

{IMPLEMENTATION}
IF i_xSetMotionPovmdEn THEN
	wMode:=i_wMotorEnMode;
	IF (i_iStationId>=0 AND i_iStationId<MAX_UNIT_NUM) THEN
		IF wMode=3 OR wMode=4 THEN
			(*iRtn:= GTD_SetMotionPovmd(1,wMode,i_iStationId);*);(*临时屏蔽|2025.08.22.134427*)
		ELSE
			iRtn:=0;
		END_IF
	ELSE
		iRtn:=-1;
	END_IF
END_IF
KS_SetMotionPovmd:=iRtn;

(* ---- KS_FB_PhaseSave.st ---- *)
(*@CES
Name=KS_FB_PhaseSave
Type=FunctionBlock
TypeGuid=6f9dac99-8de1-4efc-8465-68ac443b7d08
Guid=d61b799b-f06c-4921-af68-2abc80af0788
HasDeclaration=True
HasImplementation=True
*)
{DECLARATION}
FUNCTION_BLOCK KS_FB_PhaseSave
(*运城制版单独保存相位方式@2024.12.25.113018+注释*)
(*2025.1.3.165653 增加了每个轴的原点信号是否获取到的检查*)
(*2025.1.13.191447 增加了可以保存和可以读取标志,对输入重新做了处理*)
VAR_INPUT
	i_xEn:BOOL;
	i_xCanSave:BOOL;(*可以保存*)
	i_xBtnSave:BOOL;(*保存按钮*)
	i_xCanRead:BOOL;(*可以读取标志*)
	i_xBtnRead:BOOL;(*读取按钮*)
	(*轴的一些参数*)
	i_iGrpAxisNum_Pu: INT;(*色组轴的数量|*)
	i_aiGrpAxisList: ARRAY [1..MAX_UNIT_NUM] OF INT;(*系内所有轴的id列表,色组部分已经按照从小到大的顺序排序了，之后的是牵引|*)
	i_pstStSysParam: POINTER TO StSysParam;
//	i_pastStPTSts: POINTER TO ARRAY [1..MAX_UNIT_NUM] OF StPTSts;(*PT运动轴的状态|*)
END_VAR
VAR_OUTPUT
	o_xEn:BOOL;
END_VAR
VAR_IN_OUT
	io_xFlag_Save:BOOL;(*2024.12.25.110101 替换为了输入输出变量@作为系统保持变量了*)
	io_xFlag_Read:BOOL;(*2024.12.25.110101 替换为了输入输出变量@作为系统保持变量了*)
END_VAR
VAR
	xFlag_Save:BOOL;
	xFlag_Read:BOOL;
	iN: INT;
	iUnitId: INT;
//	pstStPTSts: POINTER TO StPTSts;(*PT运动轴的状态|*)
	fbTrig_Save:R_TRIG;
	fbTrig_Read:R_TRIG;
END_VAR
{IMPLEMENTATION}
IF i_xEn AND
	i_pstStSysParam<>0 THEN
	(*保存相位*)
	(*保存按钮操作*)
	IF i_xCanSave THEN
		fbTrig_Save(CLK:=i_xBtnSave);
		IF fbTrig_Save.Q THEN
			xFlag_Save:=TRUE;
		END_IF
	ELSE
		fbTrig_Save(CLK:=FALSE);
		xFlag_Save:=FALSE;
	END_IF

	IF xFlag_Save THEN
		FOR iN:=1 TO i_iGrpAxisNum_Pu BY 1DO
			iUnitId:=i_aiGrpAxisList[iN];
			IF i_pstStSysParam^.astStUnitParam_UnSave[iUnitId].wVirTual_Sts.12=1 THEN(*获取到了原点位置*)
				i_pstStSysParam^.astStUnitParam_Save[iUnitId].iPhase_Locating:=KS_GetPhaseValue(i_pstStSysParam^.astStUnitParam_UnSave[iUnitId].wVirTual_Cnt,gc_iVirEncPPR);
				IF iN=i_iGrpAxisNum_Pu THEN(*所有轴都没问题了*)
					xFlag_Save:=FALSE;(*复位标志*)
					io_xFlag_Save:=TRUE;(*保存成功*)
				END_IF
			ELSE(*有一个没获取到就退出*)
				xFlag_Save:=FALSE;
				io_xFlag_Save:=FALSE;
				EXIT;
			END_IF
		END_FOR
	END_IF

	(*读取相位*)
	(*读取按钮操作*)
	IF i_xCanRead THEN
		fbTrig_Read(CLK:=i_xBtnRead);
		IF fbTrig_Read.Q THEN
			io_xFlag_Read:=TRUE(*io_xFlag_Save*);(*保存成功了,就可以输出读取标志了|该变量由KS_FB_PreRegisterEtc清除*)
		END_IF
	ELSE(*不能读取就退出*)
		io_xFlag_Read:=FALSE;
		fbTrig_Read(CLK:=FALSE);
	END_IF
ELSE
	fbTrig_Save(CLK:=FALSE);
	fbTrig_Read(CLK:=FALSE);
	io_xFlag_Read:=FALSE;
	io_xFlag_Save:=FALSE;
	xFlag_Read:=FALSE;
	xFlag_Save:=FALSE;
END_IF

(* ---- KS_FB_PreRegisterCorrDeal.st ---- *)
(*@CES
Name=KS_FB_PreRegisterCorrDeal
Type=FunctionBlock
TypeGuid=6f9dac99-8de1-4efc-8465-68ac443b7d08
Guid=d37d2e52-5732-4406-aa4d-f154e1ea1a79
HasDeclaration=True
HasImplementation=True
*)
{DECLARATION}
FUNCTION_BLOCK KS_FB_PreRegisterCorrDeal
(*2024.01.15.151146 将总的调整量修改为接口*)
VAR_INPUT
	i_xEn:BOOL;(*功能块使能*)
	i_iGrpId:int;(*系号*)
	i_iGrpAxisNum_Pu: INT; (*色组轴数量*)
	i_paiGrpAxisList: POINTER TO ARRAY [1..MAX_UNIT_NUM] OF INT; (*系内所有轴的列表*)
	i_pstStSysParam: POINTER TO StSysParam;
	i_palrTotalAdjustVal_V:POINTER TO ARRAY [1..MAX_UNIT_NUM] OF LREAL;(*套色总的调整量|mm*)
END_VAR
VAR_OUTPUT
	o_xEn:BOOL;(**)
END_VAR
VAR
	alrTotalCorrectVal: ARRAY [1..MAX_UNIT_NUM] OF LREAL;
	fbTrig_PreRegister_end: R_TRIG;
	xFlag_AutoGetCorr: BOOL;
	xFlag_PringBak: BOOL;(*上个周期的印刷标志*)
END_VAR
{IMPLEMENTATION}
IF (i_iGrpId=1 OR i_iGrpId=2) AND
	i_pstStSysParam<>0 AND
	i_paiGrpAxisList<>0 AND
	i_palrTotalAdjustVal_V<>0 THEN(*2024.01.15.151230*)
	IF i_xEn THEN

		fbTrig_PreRegister_end(CLK:=i_pstStSysParam^.astStGrpParam_UnSave[i_iGrpId].xFlag_PreRegister_end);
		IF fbTrig_PreRegister_end.Q THEN(*预套准完成，置位自动获取修正量标志|*)
			xFlag_AutoGetCorr:=TRUE;
		END_IF

		IF xFlag_AutoGetCorr THEN
			IF xFlag_PringBak AND NOT i_pstStSysParam^.astStGrpParam_UnSave[i_iGrpId].xFlag_Print THEN(*退出印刷状态*)
				(*复位自动获取标志*)
				xFlag_AutoGetCorr:=FALSE;
				(*置位确认标志|用于界面显示*)
				g_axCorrectConfirmBtnDisplay[i_iGrpId]:=TRUE;
			END_IF
		END_IF
		xFlag_PringBak:=i_pstStSysParam^.astStGrpParam_UnSave[i_iGrpId].xFlag_Print;

		IF g_axPreRegisterCorrConfirm[i_iGrpId] THEN(*修正量确认按钮按下*)
			g_axCorrectConfirmBtnDisplay[i_iGrpId]:=FALSE;
		END_IF

		KS_GetCorrect_PreRegister_Auto(
			xFlag_AutoGetCorr(*i_xAutoGetCorr*),
			ADR(g_axPreRegisterCorrConfirm[i_iGrpId])(*i_pxWrPreRegisterCorr*),
			i_iGrpAxisNum_Pu(*i_iGrpAxisNum_Pu*),
			i_paiGrpAxisList(*i_paiGrpAxisList*),
			i_pstStSysParam,
			i_iGrpId,
			ADR(alrTotalCorrectVal)(*i_palrTotalCorrectVal*),
			i_palrTotalAdjustVal_V(*i_palrTotalAdjustVal_V*));
	ELSE
		xFlag_AutoGetCorr:=FALSE;
		g_axCorrectConfirmBtnDisplay[i_iGrpId]:=FALSE;
		g_axPreRegisterCorrConfirm[i_iGrpId]:=FALSE;
	END_IF
END_IF
o_xEn:=i_xEn;

(* ---- KS_FB_ProcPhaseOptReq.st ---- *)
(*@CES
Name=KS_FB_ProcPhaseOptReq
Type=FunctionBlock
TypeGuid=6f9dac99-8de1-4efc-8465-68ac443b7d08
Guid=6268291a-1193-49d9-aade-964d423980f4
HasDeclaration=True
HasImplementation=True
*)
{DECLARATION}
FUNCTION_BLOCK KS_FB_ProcPhaseOptReq (*0成功/-1参数错误|*)
(*2023.10.16.161503  处理轴的初始相位获取功能@mark线和键槽有固定相位|预套准的时候不需要手工对mark线*)
(*2023.10.17.085925|+i_xFlag_LinkageAtleast接口 *)
(*2025.1.12.171334 增加在不使能byAxisInitPhaseTypeWhenPreRegister(=1)时预套准记录mark线位置实现*)
(*2025.1.13.191531 新增加的固定相位功能在其他预套使能条件上增加*)
VAR_INPUT
	i_xEn:BOOL;
	i_iGrpId: INT;
	i_iGrpAxisNum_Pu: INT;(*色组轴的数量|*)
	i_aiGrpAxisList: ARRAY [1..MAX_UNIT_NUM] OF INT;(*系内所有轴的id列表,色组部分已经按照从小到大的顺序排序了，之后的是牵引|*)
	i_pstStSysParam: POINTER TO StSysParam;
//	i_pastStPTSts: POINTER TO ARRAY [1..MAX_UNIT_NUM] OF StPTSts;(*PT运动轴的状态|*)
	i_pxFlag_CphCommonVir: POINTER TO BOOL;
	i_pxCphaseRestore: POINTER TO BOOL;
	i_pxFlag_CphCommonVir_end: POINTER TO BOOL;
	i_pxCphaseRestore_end: POINTER TO BOOL;
	i_xFlag_LinkageAtleast1:BOOL;(*2023.10.17.085835  至少联动一色标志|改标志有效的时候预套准相关按钮不能有效*)
	(*2025.1.3.164800+目前只有运城制版使用*)
	i_xFixedPhaseSave:BOOL;(*固定的相位保存@外部需要清除*)
	i_xFixedPhaseRead:BOOL;(*固定的相位读取@外部需要清除*)
END_VAR
VAR_OUTPUT
	o_xEn:BOOL;
	o_iErrCode:INT;
END_VAR
VAR
	iN: INT;
	iUnitId: INT;
	(*2023.10.16.155940 初始原点位置保存标志*)
	xFlag_SaveAllData: BOOL;
	xFlag_SaveProtionData: BOOL;
	xBtn_InitPhaseHmiDis: BOOL;(*界面显示按钮*)
	xFlag_Enable: BOOL;(*一些运动的使能标志*)
	fbKS_FB_PhaseSave: KS_FB_PhaseSave;(*固定相位保存|2024.9.6.213537*)
	(*增加预套准标志沿@2025.1.12.170825*)
	fbRtrig_xFlag_PreRegister: R_TRIG;
	xFlag_CanSaveMarkPos:BOOL;(*可以记录标记位置标志*)
	byAxisInitPhaseTypeWhenPreRegister: BYTE;(*使能修改为了临时变量*)
END_VAR
{IMPLEMENTATION}
IF (i_iGrpAxisNum_Pu>=1 AND i_iGrpAxisNum_Pu<=MAX_UNIT_NUM) AND(*色组数量有效|*)
	i_pstStSysParam<>0 AND(*参数地址有效|*)
//	i_pastStPTSts<>0 AND
	i_pxFlag_CphCommonVir<>0 AND
	i_pxCphaseRestore<>0 AND
	i_pxFlag_CphCommonVir_end<>0 AND
	i_pxCphaseRestore_end<>0 THEN(*轴PT状态有效|*)
	(*判断读取绝对位置完成标志|2019.03.05.093558|niu.j*)
	FOR iN:=1 TO i_iGrpAxisNum_Pu BY 1 DO
		iUnitId:= i_aiGrpAxisList[iN];
		IF i_pstStSysParam^.astStUnitParam_Save[iUnitId].xLinkage THEN
			IF i_pstStSysParam^.astStUnitParam_UnSave[iUnitId].wVirTual_Sts.12=1 THEN
				i_pstStSysParam^.astStGrpParam_UnSave[i_iGrpId].xFlag_Home_end:= TRUE;
			ELSIF i_pstStSysParam^.astStUnitParam_UnSave[iUnitId].wVirTual_Sts.12<>1 THEN
				i_pstStSysParam^.astStGrpParam_UnSave[i_iGrpId].xFlag_Home_end:= FALSE;
				EXIT;
			END_IF
		END_IF
	END_FOR

	(*2023.10.16.161034|轴初始相位写入功能*)
	IF i_pstStSysParam^.astStGrpParam_Save[i_iGrpId].byAxisInitPhaseTypeWhenPreRegister>1 THEN(*非法值处理*)
		i_pstStSysParam^.astStGrpParam_Save[i_iGrpId].byAxisInitPhaseTypeWhenPreRegister:=0;
	END_IF

	(*********************START****************************************************)
	(*2025.1.12.170519 增加在预套准开始的时候记录mark线位置*)
	(*不用预套自动恢复mark线功能时*)
	xFlag_CanSaveMarkPos:=FALSE;
	byAxisInitPhaseTypeWhenPreRegister:=0;
	IF i_pstStSysParam^.astStGrpParam_Save[i_iGrpId].byAxisInitPhaseTypeWhenPreRegister=0 THEN
		fbRtrig_xFlag_PreRegister(CLK:=i_pstStSysParam^.astStGrpParam_UnSave[i_iGrpId].xFlag_PreRegister);
		(*刚进入预套准@触发记录mark线功能*)
		IF fbRtrig_xFlag_PreRegister.Q AND NOT i_pstStSysParam^.astStGrpParam_Save[i_iGrpId].xPreRegisterAxisId_Manu THEN
			i_pstStSysParam^.astStGrpParam_UnSave[i_iGrpId].xBtn_SaveAllData:=TRUE;
			xFlag_CanSaveMarkPos:=TRUE;
			byAxisInitPhaseTypeWhenPreRegister:=1;
		END_IF
	ELSE(*mark线和键槽固定相位时标志处理*)
		fbRtrig_xFlag_PreRegister(CLK:=FALSE);
		xFlag_CanSaveMarkPos:=(i_pstStSysParam^.astStGrpParam_UnSave[i_iGrpId].xFlag_Stop OR i_pstStSysParam^.astStGrpParam_UnSave[i_iGrpId].xFlag_EStop)AND(*急停或者停止都可以存储*)
						i_pstStSysParam^.astStGrpParam_UnSave[i_iGrpId].xFlag_Home_end AND(*所有联动轴已经有z脉冲了*)
						NOT i_pstStSysParam^.astStGrpParam_UnSave[i_iGrpId].xFlag_AllInchRun AND(*整机单运行*)
						NOT i_pstStSysParam^.astStGrpParam_UnSave[i_iGrpId].xFlag_Home AND(*读取装版相位*)
						NOT i_pstStSysParam^.astStGrpParam_UnSave[i_iGrpId].xFlag_PreRegister AND(*预套准*)
						NOT i_pstStSysParam^.astStGrpParam_UnSave[i_iGrpId].xFlag_PhaseRestore(*相位恢复*);

		byAxisInitPhaseTypeWhenPreRegister:=i_pstStSysParam^.astStGrpParam_Save[i_iGrpId].byAxisInitPhaseTypeWhenPreRegister;
	END_IF
	(******************END*******************************************************)

	KS_GetAxisInitPhaseWhenPreRegister(
		byAxisInitPhaseTypeWhenPreRegister(*i_byAxisInitPhaseTypeWhenPreRegister*),
		xFlag_CanSaveMarkPos(*i_xFlag_CanSaveData*),
		i_pstStSysParam^.astStGrpParam_UnSave[i_iGrpId].xBtn_SaveAllData(*i_xBtn_SaveAllData*),
		i_pstStSysParam^.astStGrpParam_UnSave[i_iGrpId].xBtn_SaveProtionData(*i_xBtn_SaveProtionData*),
		i_pstStSysParam^.astStGrpParam_UnSave[i_iGrpId].xBtn_SaveCancel(*i_xBtn_SaveCancel*),
		xBtn_InitPhaseHmiDis(*i_xBtn_DisHmi*),
		i_iGrpAxisNum_Pu(*i_iGrpAxisNum_Pu*),
		i_aiGrpAxisList(*i_aiGrpAxisList*),
		i_pstStSysParam,
//		i_pastStPTSts(*i_pastStPTSts*),
		ADR(i_pstStSysParam^.astStGrpParam_UnSave[i_iGrpId].xFlag_AxisInitPhaseHmiDis)(*i_pxInitPhaseHmiSts*),
		ADR(xFlag_SaveAllData)(*i_pxFlag_SaveAll*),
		ADR(xFlag_SaveProtionData)(*i_pxFlag_SaveProtion*));
		(*按钮清除*)
		i_pstStSysParam^.astStGrpParam_UnSave[i_iGrpId].xBtn_SaveAllData:=FALSE;
		i_pstStSysParam^.astStGrpParam_UnSave[i_iGrpId].xBtn_SaveProtionData:=FALSE;
		i_pstStSysParam^.astStGrpParam_UnSave[i_iGrpId].xBtn_SaveCancel:=FALSE;
		xBtn_InitPhaseHmiDis:=FALSE;
	(*2023.10.16.161034|轴初始相位写入功能*)

		(*2024.6.22.164252|固定相位保存*)
		fbKS_FB_PhaseSave(
			i_xEn:= TRUE,
			i_xCanSave:= (i_pstStSysParam^.astStGrpParam_UnSave[i_iGrpId].xFlag_Stop OR i_pstStSysParam^.astStGrpParam_UnSave[i_iGrpId].xFlag_EStop)AND(*急停或者停止都可以存储*)
						i_pstStSysParam^.astStGrpParam_UnSave[i_iGrpId].xFlag_Home_end AND(*所有联动轴已经有z脉冲了*)
						NOT i_pstStSysParam^.astStGrpParam_UnSave[i_iGrpId].xFlag_AllInchRun AND(*整机单运行*)
						NOT i_pstStSysParam^.astStGrpParam_UnSave[i_iGrpId].xFlag_Home AND
						NOT i_pstStSysParam^.astStGrpParam_UnSave[i_iGrpId].xFlag_PreRegister AND
						NOT i_pstStSysParam^.astStGrpParam_UnSave[i_iGrpId].xFlag_PhaseRestore,(*读取装版相位*)
			i_xBtnSave:= i_xFixedPhaseSave,
			i_xCanRead:=(i_pstStSysParam^.astStGrpParam_UnSave[i_iGrpId].xFlag_Stop)AND(*停止可以读取*)
						i_pstStSysParam^.astStGrpParam_UnSave[i_iGrpId].xFlag_Home_end AND(*所有联动轴已经有z脉冲了*)
						NOT i_pstStSysParam^.astStGrpParam_UnSave[i_iGrpId].xFlag_AllInchRun AND(*整机单运行*)
						NOT i_pstStSysParam^.astStGrpParam_UnSave[i_iGrpId].xFlag_Home AND
						NOT i_pstStSysParam^.astStGrpParam_UnSave[i_iGrpId].xFlag_PreRegister AND
						NOT i_pstStSysParam^.astStGrpParam_UnSave[i_iGrpId].xFlag_PhaseRestore,(*2025.1.13.180858+*)
			i_xBtnRead:= i_xFixedPhaseRead,
			i_iGrpAxisNum_Pu:= i_iGrpAxisNum_Pu,
			i_aiGrpAxisList:= i_aiGrpAxisList,
			i_pstStSysParam:= i_pstStSysParam,
	//		i_pastStPTSts:= i_pastStPTSts,
			io_xFlag_Save:=i_pstStSysParam^.astStGrpParam_UnSave[i_iGrpId].xFlag_PhaseSave,(*2024.12.25.110424+*)
			io_xFlag_Read:= i_pstStSysParam^.astStGrpParam_UnSave[i_iGrpId].xFlag_PhaseRead,(*2024.12.25.112509*)
			o_xEn=>);

	IF i_pstStSysParam^.astStGrpParam_UnSave[i_iGrpId].xBtn_Home THEN(*绝对位置确认/回原点|*)
		(*2023.10.17.090304*)
		xFlag_Enable:=i_pstStSysParam^.astStGrpParam_UnSave[i_iGrpId].xFlag_Stop AND
			(NOT i_pstStSysParam^.astStGrpParam_UnSave[i_iGrpId].xFlag_AllInchRun) AND
			(NOT i_pstStSysParam^.astStGrpParam_UnSave[i_iGrpId].xFlag_Estop) AND
			(NOT i_pstStSysParam^.astStGrpParam_UnSave[i_iGrpId].xFlag_EStoping) AND

			i_xFlag_LinkageAtleast1;

		IF i_pstStSysParam^.astStGrpParam_UnSave[i_iGrpId].xFlag_Home OR
			i_pstStSysParam^.astStGrpParam_UnSave[i_iGrpId].xFlag_PreRegister OR
			i_pstStSysParam^.astStGrpParam_UnSave[i_iGrpId].xFlag_PhaseRestore OR
			i_pstStSysParam^.astStGrpParam_UnSave[i_iGrpId].xFlag_PhaseRead THEN;
		ELSIF xFlag_Enable THEN(*2023.10.17.090009*)

			i_pstStSysParam^.astStGrpParam_UnSave[i_iGrpId].xFlag_Home:= TRUE;
		END_IF
		i_pstStSysParam^.astStGrpParam_UnSave[i_iGrpId].xBtn_Home:= FALSE;

		IF g_iPrewrkSubPageId=1 THEN(*2023.10.16.161006@处于纵向预套准界面点击读取装版相位才显示*)
			xBtn_InitPhaseHmiDis:=TRUE;(*2023.10.16.161006|显示初始相位保存界面*)
		END_IF

	ELSIF i_pstStSysParam^.astStGrpParam_UnSave[i_iGrpId].xBtn_ConfirmPreRegHomePos THEN(*保存装版位|*)
		i_pstStSysParam^.astStGrpParam_UnSave[i_iGrpId].xFlag_ConfirmPreRegHomePos:= TRUE;
		i_pstStSysParam^.astStGrpParam_UnSave[i_iGrpId].xFlag_ConfirmPreRegHomePos_ing:= TRUE;
		i_pstStSysParam^.astStGrpParam_UnSave[i_iGrpId].xFlag_ConfirmPreRegHomePos_end:= FALSE;

		IF i_pstStSysParam^.astStGrpParam_UnSave[i_iGrpId].xFlag_Home_end THEN (*回原点完成*)
			FOR iN:=1 TO i_iGrpAxisNum_Pu BY 1 DO
				iUnitId:= i_aiGrpAxisList[iN];

				IF i_pstStSysParam^.astStUnitParam_Save[iUnitId].xLinkage THEN
					(*2023.6.28.113335 更新*)
					i_pstStSysParam^.astStUnitParam_UnSave[iUnitId].iPhase_InstallPlate:=KS_GetPhaseValue(i_pstStSysParam^.astStUnitParam_UnSave[iUnitId].wVirTual_Cnt,gc_iVirEncPPR);

				END_IF
			END_FOR

			i_pstStSysParam^.astStGrpParam_UnSave[i_iGrpId].xFlag_ConfirmPreRegHomePos_end:= TRUE;
		END_IF

		i_pstStSysParam^.astStGrpParam_UnSave[i_iGrpId].xFlag_ConfirmPreRegHomePos_ing:= FALSE;
		i_pstStSysParam^.astStGrpParam_UnSave[i_iGrpId].xFlag_ConfirmPreRegHomePos:= FALSE;

		i_pstStSysParam^.astStGrpParam_UnSave[i_iGrpId].xBtn_ConfirmPreRegHomePos:= FALSE;
	ELSIF i_pstStSysParam^.astStGrpParam_UnSave[i_iGrpId].xBtn_PreRegister THEN(*纵向预套准|*)
		IF i_pstStSysParam^.astStGrpParam_UnSave[i_iGrpId].xFlag_Home OR
			i_pstStSysParam^.astStGrpParam_UnSave[i_iGrpId].xFlag_PreRegister OR
			i_pstStSysParam^.astStGrpParam_UnSave[i_iGrpId].xFlag_PhaseRestore OR
			i_pstStSysParam^.astStGrpParam_UnSave[i_iGrpId].xFlag_PhaseRead THEN
			;
		ELSIF i_pstStSysParam^.astStGrpParam_UnSave[i_iGrpId].xFlag_Stop AND
			(NOT i_pstStSysParam^.astStGrpParam_UnSave[i_iGrpId].xFlag_AllInchRun) AND
			(NOT i_pstStSysParam^.astStGrpParam_UnSave[i_iGrpId].xFlag_Estop) AND
			(NOT i_pstStSysParam^.astStGrpParam_UnSave[i_iGrpId].xFlag_EStoping) AND
			i_pstStSysParam^.astStGrpParam_UnSave[i_iGrpId].xFlag_Home_end AND
			(i_xFlag_LinkageAtleast1 ) THEN(*2023.10.17.090009*)
			;
			i_pstStSysParam^.astStGrpParam_UnSave[i_iGrpId].xFlag_PreRegister:= TRUE;
		END_IF
		i_pstStSysParam^.astStGrpParam_UnSave[i_iGrpId].xBtn_PreRegister:= FALSE;
	ELSIF g_xLoadRecipe_End THEN(*相位恢复|*)
		IF i_pstStSysParam^.astStGrpParam_UnSave[i_iGrpId].xFlag_Home OR
			i_pstStSysParam^.astStGrpParam_UnSave[i_iGrpId].xFlag_PreRegister OR
			i_pstStSysParam^.astStGrpParam_UnSave[i_iGrpId].xFlag_PhaseRestore OR
			i_pstStSysParam^.astStGrpParam_UnSave[i_iGrpId].xFlag_PhaseRead THEN
			;
		ELSIF i_pstStSysParam^.astStGrpParam_UnSave[i_iGrpId].xFlag_Stop AND
			(NOT i_pstStSysParam^.astStGrpParam_UnSave[i_iGrpId].xFlag_AllInchRun) AND
			(NOT i_pstStSysParam^.astStGrpParam_UnSave[i_iGrpId].xFlag_Estop) AND
			(NOT i_pstStSysParam^.astStGrpParam_UnSave[i_iGrpId].xFlag_EStoping) AND
			i_pstStSysParam^.astStGrpParam_UnSave[i_iGrpId].xFlag_Home_end AND
			(i_xFlag_LinkageAtleast1 ) THEN(*2023.10.17.090009*)
			;
			i_pstStSysParam^.astStGrpParam_UnSave[i_iGrpId].xFlag_PhaseRestore:= TRUE;

		END_IF
		g_xLoadRecipe_End:= FALSE;
	ELSIF i_pstStSysParam^.astStGrpParam_UnSave[i_iGrpId].xBtn_PhaseSave THEN(*相位保存|*)
		i_pstStSysParam^.astStGrpParam_UnSave[i_iGrpId].xBtn_PhaseSave:= FALSE;

		FOR iN:=1 TO i_iGrpAxisNum_Pu BY 1 DO
			iUnitId:= i_aiGrpAxisList[iN];
			(*2021.9.18.113751 增加相位保存时候变量初始化*)
			i_pstStSysParam^.astStUnitParam_UnSave[iUnitId].iPhase_RegisterOk:=0;
			IF i_pstStSysParam^.astStUnitParam_Save[iUnitId].xLinkage THEN
				(*2023.6.28.113526 更新*)
				i_pstStSysParam^.astStUnitParam_UnSave[iUnitId].iPhase_RegisterOk:=KS_GetPhaseValue(i_pstStSysParam^.astStUnitParam_UnSave[iUnitId].wVirTual_Cnt,gc_iVirEncPPR);

				(*非负保护|2021.10.25.154529*)
				IF i_pstStSysParam^.astStUnitParam_UnSave[iUnitId].iPhase_RegisterOk < 0 THEN
					i_pstStSysParam^.astStUnitParam_UnSave[iUnitId].iPhase_RegisterOk:=0;
				END_IF
			END_IF
		END_FOR
		(*2018.11.5.132513|相位保存完成，直接进去配方写入流程*)
		g_xReqSaveRecipe:=TRUE; (*写入配方使能*)

(*2019.07.27.164458|niu.j|通用配方逻辑处理*)
	ELSIF g_xReqSaveCphRecipe THEN
		g_xReqSaveCphRecipe:=FALSE;
		FOR iN:=1 TO i_iGrpAxisNum_Pu BY 1 DO
			iUnitId:= i_aiGrpAxisList[iN];

			(*2021.9.18.113751 增加相位保存时候变量初始化*)
			i_pstStSysParam^.astStUnitParam_Save[iUnitId].iPhase_RegisterOk:=0;
			i_pstStSysParam^.astStUnitParam_Save[iUnitId].iPhase_FinalUsed:=0;
			IF i_pstStSysParam^.astStUnitParam_Save[iUnitId].xLinkage THEN
				(*2023.6.28.113822 更新*)
				i_pstStSysParam^.astStUnitParam_Save[iUnitId].iPhase_RegisterOk:=KS_GetPhaseValue(i_pstStSysParam^.astStUnitParam_UnSave[iUnitId].wVirTual_Cnt,gc_iVirEncPPR);

				i_pstStSysParam^.astStUnitParam_Save[iUnitId].iPhase_FinalUsed:= i_pstStSysParam^.astStUnitParam_Save[iUnitId].iPhase_RegisterOk-i_pstStSysParam^.astStUnitParam_Save[iUnitId].iPhase_InstallPlate;

				WHILE i_pstStSysParam^.astStUnitParam_Save[iUnitId].iPhase_FinalUsed<0 DO
					i_pstStSysParam^.astStUnitParam_Save[iUnitId].iPhase_FinalUsed:= i_pstStSysParam^.astStUnitParam_Save[iUnitId].iPhase_FinalUsed+gc_iVirEncPPR;
				END_WHILE

				WHILE i_pstStSysParam^.astStUnitParam_Save[iUnitId].iPhase_FinalUsed>=gc_iVirEncPPR DO (* 2021.7.1.104815/ *)
					i_pstStSysParam^.astStUnitParam_Save[iUnitId].iPhase_FinalUsed:= i_pstStSysParam^.astStUnitParam_Save[iUnitId].iPhase_FinalUsed-gc_iVirEncPPR;
				END_WHILE
			END_IF
		END_FOR
		(*2018.11.5.132513|相位保存完成，直接进去配方写入流程*)

(*初始相位保存*)
	ELSIF g_xReqSaveCphCommonVir THEN
		IF i_pstStSysParam^.astStGrpParam_UnSave[i_iGrpId].xFlag_Home OR
			i_pstStSysParam^.astStGrpParam_UnSave[i_iGrpId].xFlag_PreRegister OR
			i_pstStSysParam^.astStGrpParam_UnSave[i_iGrpId].xFlag_PhaseRestore OR
			i_pxFlag_CphCommonVir^ THEN
			;
		ELSIF i_pstStSysParam^.astStGrpParam_UnSave[i_iGrpId].xFlag_Stop AND
			(NOT i_pstStSysParam^.astStGrpParam_UnSave[i_iGrpId].xFlag_AllInchRun) AND
			(NOT i_pstStSysParam^.astStGrpParam_UnSave[i_iGrpId].xFlag_Estop) AND
			(NOT i_pstStSysParam^.astStGrpParam_UnSave[i_iGrpId].xFlag_EStoping) AND
			(NOT i_pxFlag_CphCommonVir^) THEN
			;
			i_pxFlag_CphCommonVir^:= TRUE;
		END_IF
		IF NOT i_pxFlag_CphCommonVir_end^ THEN
			;
		ELSE
			FOR iN:=1 TO i_iGrpAxisNum_Pu BY 1 DO
				iUnitId:= i_aiGrpAxisList[iN];

				IF i_pstStSysParam^.astStUnitParam_Save[iUnitId].xLinkage THEN
					(*2023.6.28.113642 更新*)
					i_pstStSysParam^.astStUnitParam_Save[iUnitId].iPhase_InstallPlate:=KS_GetPhaseValue(i_pstStSysParam^.astStUnitParam_UnSave[iUnitId].wVirTual_Cnt,gc_iVirEncPPR);
				END_IF
			END_FOR
			g_xReqSaveCphCommonVir:= FALSE;
		END_IF

	ELSIF g_xLoadCphRecipe_End THEN
		IF i_pstStSysParam^.astStGrpParam_UnSave[i_iGrpId].xFlag_Home OR
			i_pstStSysParam^.astStGrpParam_UnSave[i_iGrpId].xFlag_PreRegister OR
			i_pstStSysParam^.astStGrpParam_UnSave[i_iGrpId].xFlag_PhaseRestore THEN
			;
		ELSIF i_pstStSysParam^.astStGrpParam_UnSave[i_iGrpId].xFlag_Stop AND
			(NOT i_pstStSysParam^.astStGrpParam_UnSave[i_iGrpId].xFlag_AllInchRun) AND
			(NOT i_pstStSysParam^.astStGrpParam_UnSave[i_iGrpId].xFlag_Estop) AND
			(NOT i_pstStSysParam^.astStGrpParam_UnSave[i_iGrpId].xFlag_EStoping) AND
			i_pxFlag_CphCommonVir_end^ THEN
			;
			i_pxCphaseRestore^:= TRUE;
		END_IF
		g_xLoadCphRecipe_End:= FALSE;
	END_IF

	o_iErrCode:= 0;
ELSE
	o_iErrCode:= -1;
END_IF
